DATA_BLOCK DB 50
VERSION : 0.1


  STRUCT
   STAT0 : DATE_AND_TIME  := DT#95-1-1-0:0:0.000;
   STAT1 : DATE_AND_TIME  := DT#95-1-1-0:0:0.000;
   STAT2 : INT ;
   STAT3 : DATE  := D#1995-1-1;
   STAT4 : TIME_OF_DAY ;
   STAT5 : INT ;
   STAT6 : BYTE ;
  END_STRUCT ;
BEGIN
   STAT0 := DT#22-2-18-16:13:36.401;
   STAT1 := DT#95-1-1-0:0:0.000;
   STAT2 := 0;
   STAT3 := D#1995-1-1;
   STAT4 := TOD#0:0:0.000;
   STAT5 := 0;
   STAT6 := B#16#0;
END_DATA_BLOCK

DATA_BLOCK DB 101
VERSION : 0.1


  STRUCT
   STAT0 : STRUCT
    STAT1 : STRUCT
     STAT2 : WORD ;
     STAT3 : WORD ;
    END_STRUCT ;
    STAT4 : STRUCT
     STAT5 : WORD ;
     STAT6 : STRUCT
      STAT7 : BOOL ;
      STAT8 : BOOL ;
      STAT9 : BOOL ;
      STAT10 : BOOL ;
      STAT11 : BOOL ;
      STAT12 : BOOL ;
      STAT13 : BOOL ;
      STAT14 : BOOL ;
      STAT15 : BOOL ;
      STAT16 : BOOL ;
      STAT17 : BOOL ;
      STAT18 : BOOL ;
      STAT19 : BOOL ;
      STAT20 : BOOL ;
      STAT21 : BOOL ;
      STAT22 : BOOL ;
     END_STRUCT ;
     STAT23 : WORD ;
     STAT24 : WORD ;
     STAT25 : WORD ;
     STAT26 : WORD ;
     STAT27 : WORD ;
     STAT28 : BYTE ;
     STAT29 : BYTE ;
    END_STRUCT ;
    STAT30 : BOOL ;
    STAT31 : BOOL ;
    STAT32 : WORD ;
    STAT33 : INT ;
   END_STRUCT ;
   STAT34 : STRUCT
    STAT35 : STRUCT
     STAT36 : WORD ;
     STAT37 : WORD ;
    END_STRUCT ;
    STAT38 : STRUCT
     STAT39 : ARRAY  [0 .. 12 ] OF STRUCT
      STAT40 : BOOL ;
      STAT41 : BOOL ;
      STAT42 : BOOL ;
      STAT43 : BOOL ;
      STAT44 : BOOL ;
      STAT45 : BOOL ;
      STAT46 : BOOL ;
      STAT47 : BOOL ;
      STAT48 : BYTE ;
      STAT49 : BYTE ;
      STAT50 : BYTE ;
     END_STRUCT ;
     STAT51 : ARRAY  [0 .. 12 ] OF STRUCT
      STAT52 : BOOL ;
      STAT53 : BOOL ;
      STAT54 : BOOL ;
      STAT55 : BOOL ;
      STAT56 : BOOL ;
      STAT57 : BOOL ;
      STAT58 : BOOL ;
      STAT59 : BOOL ;
      STAT60 : BYTE ;
      STAT61 : BYTE ;
      STAT62 : BYTE ;
     END_STRUCT ;
    END_STRUCT ;
    STAT63 : BOOL ;
    STAT64 : BOOL ;
    STAT65 : WORD ;
    STAT66 : INT ;
   END_STRUCT ;
   STAT67 : STRUCT
    STAT68 : STRUCT
     STAT69 : WORD ;
     STAT70 : WORD ;
    END_STRUCT ;
    STAT71 : STRUCT
     STAT72 : WORD ;
     STAT73 : WORD ;
     STAT74 : WORD ;
     STAT75 : WORD ;
     STAT76 : WORD ;
     STAT77 : WORD ;
     STAT78 : WORD ;
     STAT79 : STRUCT
      STAT80 : BOOL ;
      STAT81 : BOOL ;
      STAT82 : BOOL ;
      STAT83 : BOOL ;
      STAT84 : BOOL ;
      STAT85 : BOOL ;
      STAT86 : BOOL ;
      STAT87 : BOOL ;
      STAT88 : BOOL ;
      STAT89 : BOOL ;
      STAT90 : BOOL ;
      STAT91 : BOOL ;
      STAT92 : BOOL ;
      STAT93 : BOOL ;
      STAT94 : BOOL ;
      STAT95 : BOOL ;
     END_STRUCT ;
    END_STRUCT ;
    STAT96 : BOOL ;
    STAT97 : BOOL ;
    STAT98 : WORD ;
    STAT99 : INT ;
   END_STRUCT ;
   STAT100 : STRUCT
    STAT101 : STRUCT
     STAT102 : WORD ;
     STAT103 : WORD ;
    END_STRUCT ;
    STAT104 : STRUCT
     STAT105 : WORD ;
     STAT106 : WORD ;
     STAT107 : WORD ;
     STAT108 : WORD ;
     STAT109 : WORD ;
     STAT110 : WORD ;
     STAT111 : WORD ;
     STAT112 : STRUCT
      STAT113 : BOOL ;
      STAT114 : BOOL ;
      STAT115 : BOOL ;
      STAT116 : BOOL ;
      STAT117 : BOOL ;
      STAT118 : BOOL ;
      STAT119 : BOOL ;
      STAT120 : BOOL ;
      STAT121 : BOOL ;
      STAT122 : BOOL ;
      STAT123 : BOOL ;
      STAT124 : BOOL ;
      STAT125 : BOOL ;
      STAT126 : BOOL ;
      STAT127 : BOOL ;
      STAT128 : BOOL ;
     END_STRUCT ;
    END_STRUCT ;
    STAT129 : BOOL ;
    STAT130 : BOOL ;
    STAT131 : WORD ;
    STAT132 : INT ;
   END_STRUCT ;
   STAT133 : STRUCT
    STAT134 : STRUCT
     STAT135 : WORD ;
     STAT136 : WORD ;
    END_STRUCT ;
    STAT137 : STRUCT
     STAT138 : WORD ;
     STAT139 : WORD ;
     STAT140 : WORD ;
     STAT141 : WORD ;
     STAT142 : WORD ;
     STAT143 : WORD ;
     STAT144 : WORD ;
     STAT145 : STRUCT
      STAT146 : BOOL ;
      STAT147 : BOOL ;
      STAT148 : BOOL ;
      STAT149 : BOOL ;
      STAT150 : BOOL ;
      STAT151 : BOOL ;
      STAT152 : BOOL ;
      STAT153 : BOOL ;
      STAT154 : BOOL ;
      STAT155 : BOOL ;
      STAT156 : BOOL ;
      STAT157 : BOOL ;
      STAT158 : BOOL ;
      STAT159 : BOOL ;
      STAT160 : BOOL ;
      STAT161 : BOOL ;
     END_STRUCT ;
    END_STRUCT ;
    STAT162 : BOOL ;
    STAT163 : BOOL ;
    STAT164 : WORD ;
    STAT165 : INT ;
   END_STRUCT ;
   STAT166 : BYTE ;
   STAT167 : BYTE ;
   STAT168 : ARRAY  [0 .. 25 ] OF STRUCT
    STAT169 : BOOL ;
    STAT170 : BOOL ;
    STAT171 : BOOL ;
    STAT172 : BOOL ;
    STAT173 : BOOL ;
    STAT174 : BOOL ;
    STAT175 : BOOL ;
    STAT176 : BOOL ;
    STAT177 : BYTE ;
    STAT178 : BYTE ;
    STAT179 : BYTE ;
   END_STRUCT ;
  END_STRUCT ;
BEGIN
   STAT0.STAT1.STAT2 := W#16#10;
   STAT0.STAT1.STAT3 := W#16#1;
   STAT0.STAT4.STAT5 := W#16#12;
   STAT0.STAT4.STAT6.STAT7 := FALSE;
   STAT0.STAT4.STAT6.STAT8 := FALSE;
   STAT0.STAT4.STAT6.STAT9 := FALSE;
   STAT0.STAT4.STAT6.STAT10 := FALSE;
   STAT0.STAT4.STAT6.STAT11 := TRUE;
   STAT0.STAT4.STAT6.STAT12 := FALSE;
   STAT0.STAT4.STAT6.STAT13 := FALSE;
   STAT0.STAT4.STAT6.STAT14 := FALSE;
   STAT0.STAT4.STAT6.STAT15 := TRUE;
   STAT0.STAT4.STAT6.STAT16 := FALSE;
   STAT0.STAT4.STAT6.STAT17 := FALSE;
   STAT0.STAT4.STAT6.STAT18 := FALSE;
   STAT0.STAT4.STAT6.STAT19 := FALSE;
   STAT0.STAT4.STAT6.STAT20 := FALSE;
   STAT0.STAT4.STAT6.STAT21 := FALSE;
   STAT0.STAT4.STAT6.STAT22 := FALSE;
   STAT0.STAT4.STAT23 := W#16#0;
   STAT0.STAT4.STAT24 := W#16#0;
   STAT0.STAT4.STAT25 := W#16#9;
   STAT0.STAT4.STAT26 := W#16#9;
   STAT0.STAT4.STAT27 := W#16#0;
   STAT0.STAT4.STAT28 := B#16#3;
   STAT0.STAT4.STAT29 := B#16#0;
   STAT0.STAT30 := TRUE;
   STAT0.STAT31 := FALSE;
   STAT0.STAT32 := W#16#0;
   STAT0.STAT33 := 0;
   STAT34.STAT35.STAT36 := W#16#4;
   STAT34.STAT35.STAT37 := W#16#18;
   STAT34.STAT38.STAT39[0].STAT40 := FALSE;
   STAT34.STAT38.STAT39[0].STAT41 := FALSE;
   STAT34.STAT38.STAT39[0].STAT42 := FALSE;
   STAT34.STAT38.STAT39[0].STAT43 := TRUE;
   STAT34.STAT38.STAT39[0].STAT44 := TRUE;
   STAT34.STAT38.STAT39[0].STAT45 := TRUE;
   STAT34.STAT38.STAT39[0].STAT46 := TRUE;
   STAT34.STAT38.STAT39[0].STAT47 := TRUE;
   STAT34.STAT38.STAT39[0].STAT48 := B#16#2;
   STAT34.STAT38.STAT39[0].STAT49 := B#16#0;
   STAT34.STAT38.STAT39[0].STAT50 := B#16#0;
   STAT34.STAT38.STAT39[1].STAT40 := FALSE;
   STAT34.STAT38.STAT39[1].STAT41 := FALSE;
   STAT34.STAT38.STAT39[1].STAT42 := FALSE;
   STAT34.STAT38.STAT39[1].STAT43 := TRUE;
   STAT34.STAT38.STAT39[1].STAT44 := TRUE;
   STAT34.STAT38.STAT39[1].STAT45 := TRUE;
   STAT34.STAT38.STAT39[1].STAT46 := TRUE;
   STAT34.STAT38.STAT39[1].STAT47 := TRUE;
   STAT34.STAT38.STAT39[1].STAT48 := B#16#3;
   STAT34.STAT38.STAT39[1].STAT49 := B#16#1;
   STAT34.STAT38.STAT39[1].STAT50 := B#16#0;
   STAT34.STAT38.STAT39[2].STAT40 := FALSE;
   STAT34.STAT38.STAT39[2].STAT41 := FALSE;
   STAT34.STAT38.STAT39[2].STAT42 := FALSE;
   STAT34.STAT38.STAT39[2].STAT43 := TRUE;
   STAT34.STAT38.STAT39[2].STAT44 := TRUE;
   STAT34.STAT38.STAT39[2].STAT45 := TRUE;
   STAT34.STAT38.STAT39[2].STAT46 := TRUE;
   STAT34.STAT38.STAT39[2].STAT47 := TRUE;
   STAT34.STAT38.STAT39[2].STAT48 := B#16#4;
   STAT34.STAT38.STAT39[2].STAT49 := B#16#1;
   STAT34.STAT38.STAT39[2].STAT50 := B#16#0;
   STAT34.STAT38.STAT39[3].STAT40 := FALSE;
   STAT34.STAT38.STAT39[3].STAT41 := FALSE;
   STAT34.STAT38.STAT39[3].STAT42 := FALSE;
   STAT34.STAT38.STAT39[3].STAT43 := TRUE;
   STAT34.STAT38.STAT39[3].STAT44 := TRUE;
   STAT34.STAT38.STAT39[3].STAT45 := TRUE;
   STAT34.STAT38.STAT39[3].STAT46 := TRUE;
   STAT34.STAT38.STAT39[3].STAT47 := TRUE;
   STAT34.STAT38.STAT39[3].STAT48 := B#16#5;
   STAT34.STAT38.STAT39[3].STAT49 := B#16#0;
   STAT34.STAT38.STAT39[3].STAT50 := B#16#0;
   STAT34.STAT38.STAT39[4].STAT40 := FALSE;
   STAT34.STAT38.STAT39[4].STAT41 := FALSE;
   STAT34.STAT38.STAT39[4].STAT42 := FALSE;
   STAT34.STAT38.STAT39[4].STAT43 := TRUE;
   STAT34.STAT38.STAT39[4].STAT44 := TRUE;
   STAT34.STAT38.STAT39[4].STAT45 := TRUE;
   STAT34.STAT38.STAT39[4].STAT46 := TRUE;
   STAT34.STAT38.STAT39[4].STAT47 := TRUE;
   STAT34.STAT38.STAT39[4].STAT48 := B#16#6;
   STAT34.STAT38.STAT39[4].STAT49 := B#16#0;
   STAT34.STAT38.STAT39[4].STAT50 := B#16#0;
   STAT34.STAT38.STAT39[5].STAT40 := FALSE;
   STAT34.STAT38.STAT39[5].STAT41 := FALSE;
   STAT34.STAT38.STAT39[5].STAT42 := FALSE;
   STAT34.STAT38.STAT39[5].STAT43 := TRUE;
   STAT34.STAT38.STAT39[5].STAT44 := TRUE;
   STAT34.STAT38.STAT39[5].STAT45 := TRUE;
   STAT34.STAT38.STAT39[5].STAT46 := TRUE;
   STAT34.STAT38.STAT39[5].STAT47 := TRUE;
   STAT34.STAT38.STAT39[5].STAT48 := B#16#B;
   STAT34.STAT38.STAT39[5].STAT49 := B#16#0;
   STAT34.STAT38.STAT39[5].STAT50 := B#16#0;
   STAT34.STAT38.STAT39[6].STAT40 := FALSE;
   STAT34.STAT38.STAT39[6].STAT41 := FALSE;
   STAT34.STAT38.STAT39[6].STAT42 := FALSE;
   STAT34.STAT38.STAT39[6].STAT43 := TRUE;
   STAT34.STAT38.STAT39[6].STAT44 := TRUE;
   STAT34.STAT38.STAT39[6].STAT45 := TRUE;
   STAT34.STAT38.STAT39[6].STAT46 := TRUE;
   STAT34.STAT38.STAT39[6].STAT47 := TRUE;
   STAT34.STAT38.STAT39[6].STAT48 := B#16#D;
   STAT34.STAT38.STAT39[6].STAT49 := B#16#0;
   STAT34.STAT38.STAT39[6].STAT50 := B#16#0;
   STAT34.STAT38.STAT39[7].STAT40 := FALSE;
   STAT34.STAT38.STAT39[7].STAT41 := FALSE;
   STAT34.STAT38.STAT39[7].STAT42 := FALSE;
   STAT34.STAT38.STAT39[7].STAT43 := TRUE;
   STAT34.STAT38.STAT39[7].STAT44 := TRUE;
   STAT34.STAT38.STAT39[7].STAT45 := TRUE;
   STAT34.STAT38.STAT39[7].STAT46 := TRUE;
   STAT34.STAT38.STAT39[7].STAT47 := TRUE;
   STAT34.STAT38.STAT39[7].STAT48 := B#16#E;
   STAT34.STAT38.STAT39[7].STAT49 := B#16#1;
   STAT34.STAT38.STAT39[7].STAT50 := B#16#0;
   STAT34.STAT38.STAT39[8].STAT40 := FALSE;
   STAT34.STAT38.STAT39[8].STAT41 := FALSE;
   STAT34.STAT38.STAT39[8].STAT42 := FALSE;
   STAT34.STAT38.STAT39[8].STAT43 := TRUE;
   STAT34.STAT38.STAT39[8].STAT44 := TRUE;
   STAT34.STAT38.STAT39[8].STAT45 := TRUE;
   STAT34.STAT38.STAT39[8].STAT46 := TRUE;
   STAT34.STAT38.STAT39[8].STAT47 := TRUE;
   STAT34.STAT38.STAT39[8].STAT48 := B#16#F;
   STAT34.STAT38.STAT39[8].STAT49 := B#16#1;
   STAT34.STAT38.STAT39[8].STAT50 := B#16#0;
   STAT34.STAT38.STAT39[9].STAT40 := FALSE;
   STAT34.STAT38.STAT39[9].STAT41 := FALSE;
   STAT34.STAT38.STAT39[9].STAT42 := FALSE;
   STAT34.STAT38.STAT39[9].STAT43 := TRUE;
   STAT34.STAT38.STAT39[9].STAT44 := TRUE;
   STAT34.STAT38.STAT39[9].STAT45 := TRUE;
   STAT34.STAT38.STAT39[9].STAT46 := TRUE;
   STAT34.STAT38.STAT39[9].STAT47 := TRUE;
   STAT34.STAT38.STAT39[9].STAT48 := B#16#10;
   STAT34.STAT38.STAT39[9].STAT49 := B#16#0;
   STAT34.STAT38.STAT39[9].STAT50 := B#16#0;
   STAT34.STAT38.STAT39[10].STAT40 := FALSE;
   STAT34.STAT38.STAT39[10].STAT41 := FALSE;
   STAT34.STAT38.STAT39[10].STAT42 := FALSE;
   STAT34.STAT38.STAT39[10].STAT43 := TRUE;
   STAT34.STAT38.STAT39[10].STAT44 := TRUE;
   STAT34.STAT38.STAT39[10].STAT45 := TRUE;
   STAT34.STAT38.STAT39[10].STAT46 := TRUE;
   STAT34.STAT38.STAT39[10].STAT47 := TRUE;
   STAT34.STAT38.STAT39[10].STAT48 := B#16#12;
   STAT34.STAT38.STAT39[10].STAT49 := B#16#0;
   STAT34.STAT38.STAT39[10].STAT50 := B#16#0;
   STAT34.STAT38.STAT39[11].STAT40 := FALSE;
   STAT34.STAT38.STAT39[11].STAT41 := FALSE;
   STAT34.STAT38.STAT39[11].STAT42 := FALSE;
   STAT34.STAT38.STAT39[11].STAT43 := TRUE;
   STAT34.STAT38.STAT39[11].STAT44 := TRUE;
   STAT34.STAT38.STAT39[11].STAT45 := TRUE;
   STAT34.STAT38.STAT39[11].STAT46 := TRUE;
   STAT34.STAT38.STAT39[11].STAT47 := TRUE;
   STAT34.STAT38.STAT39[11].STAT48 := B#16#13;
   STAT34.STAT38.STAT39[11].STAT49 := B#16#0;
   STAT34.STAT38.STAT39[11].STAT50 := B#16#0;
   STAT34.STAT38.STAT39[12].STAT40 := TRUE;
   STAT34.STAT38.STAT39[12].STAT41 := FALSE;
   STAT34.STAT38.STAT39[12].STAT42 := FALSE;
   STAT34.STAT38.STAT39[12].STAT43 := FALSE;
   STAT34.STAT38.STAT39[12].STAT44 := TRUE;
   STAT34.STAT38.STAT39[12].STAT45 := TRUE;
   STAT34.STAT38.STAT39[12].STAT46 := TRUE;
   STAT34.STAT38.STAT39[12].STAT47 := TRUE;
   STAT34.STAT38.STAT39[12].STAT48 := B#16#2;
   STAT34.STAT38.STAT39[12].STAT49 := B#16#0;
   STAT34.STAT38.STAT39[12].STAT50 := B#16#0;
   STAT34.STAT38.STAT51[0].STAT52 := TRUE;
   STAT34.STAT38.STAT51[0].STAT53 := FALSE;
   STAT34.STAT38.STAT51[0].STAT54 := FALSE;
   STAT34.STAT38.STAT51[0].STAT55 := FALSE;
   STAT34.STAT38.STAT51[0].STAT56 := TRUE;
   STAT34.STAT38.STAT51[0].STAT57 := TRUE;
   STAT34.STAT38.STAT51[0].STAT58 := TRUE;
   STAT34.STAT38.STAT51[0].STAT59 := TRUE;
   STAT34.STAT38.STAT51[0].STAT60 := B#16#3;
   STAT34.STAT38.STAT51[0].STAT61 := B#16#1;
   STAT34.STAT38.STAT51[0].STAT62 := B#16#0;
   STAT34.STAT38.STAT51[1].STAT52 := TRUE;
   STAT34.STAT38.STAT51[1].STAT53 := FALSE;
   STAT34.STAT38.STAT51[1].STAT54 := FALSE;
   STAT34.STAT38.STAT51[1].STAT55 := FALSE;
   STAT34.STAT38.STAT51[1].STAT56 := TRUE;
   STAT34.STAT38.STAT51[1].STAT57 := TRUE;
   STAT34.STAT38.STAT51[1].STAT58 := TRUE;
   STAT34.STAT38.STAT51[1].STAT59 := TRUE;
   STAT34.STAT38.STAT51[1].STAT60 := B#16#4;
   STAT34.STAT38.STAT51[1].STAT61 := B#16#1;
   STAT34.STAT38.STAT51[1].STAT62 := B#16#0;
   STAT34.STAT38.STAT51[2].STAT52 := TRUE;
   STAT34.STAT38.STAT51[2].STAT53 := FALSE;
   STAT34.STAT38.STAT51[2].STAT54 := FALSE;
   STAT34.STAT38.STAT51[2].STAT55 := FALSE;
   STAT34.STAT38.STAT51[2].STAT56 := TRUE;
   STAT34.STAT38.STAT51[2].STAT57 := TRUE;
   STAT34.STAT38.STAT51[2].STAT58 := TRUE;
   STAT34.STAT38.STAT51[2].STAT59 := TRUE;
   STAT34.STAT38.STAT51[2].STAT60 := B#16#5;
   STAT34.STAT38.STAT51[2].STAT61 := B#16#0;
   STAT34.STAT38.STAT51[2].STAT62 := B#16#0;
   STAT34.STAT38.STAT51[3].STAT52 := TRUE;
   STAT34.STAT38.STAT51[3].STAT53 := FALSE;
   STAT34.STAT38.STAT51[3].STAT54 := FALSE;
   STAT34.STAT38.STAT51[3].STAT55 := FALSE;
   STAT34.STAT38.STAT51[3].STAT56 := TRUE;
   STAT34.STAT38.STAT51[3].STAT57 := TRUE;
   STAT34.STAT38.STAT51[3].STAT58 := TRUE;
   STAT34.STAT38.STAT51[3].STAT59 := TRUE;
   STAT34.STAT38.STAT51[3].STAT60 := B#16#6;
   STAT34.STAT38.STAT51[3].STAT61 := B#16#0;
   STAT34.STAT38.STAT51[3].STAT62 := B#16#0;
   STAT34.STAT38.STAT51[4].STAT52 := TRUE;
   STAT34.STAT38.STAT51[4].STAT53 := FALSE;
   STAT34.STAT38.STAT51[4].STAT54 := FALSE;
   STAT34.STAT38.STAT51[4].STAT55 := FALSE;
   STAT34.STAT38.STAT51[4].STAT56 := TRUE;
   STAT34.STAT38.STAT51[4].STAT57 := TRUE;
   STAT34.STAT38.STAT51[4].STAT58 := TRUE;
   STAT34.STAT38.STAT51[4].STAT59 := TRUE;
   STAT34.STAT38.STAT51[4].STAT60 := B#16#B;
   STAT34.STAT38.STAT51[4].STAT61 := B#16#0;
   STAT34.STAT38.STAT51[4].STAT62 := B#16#0;
   STAT34.STAT38.STAT51[5].STAT52 := TRUE;
   STAT34.STAT38.STAT51[5].STAT53 := FALSE;
   STAT34.STAT38.STAT51[5].STAT54 := FALSE;
   STAT34.STAT38.STAT51[5].STAT55 := FALSE;
   STAT34.STAT38.STAT51[5].STAT56 := TRUE;
   STAT34.STAT38.STAT51[5].STAT57 := TRUE;
   STAT34.STAT38.STAT51[5].STAT58 := TRUE;
   STAT34.STAT38.STAT51[5].STAT59 := TRUE;
   STAT34.STAT38.STAT51[5].STAT60 := B#16#D;
   STAT34.STAT38.STAT51[5].STAT61 := B#16#0;
   STAT34.STAT38.STAT51[5].STAT62 := B#16#0;
   STAT34.STAT38.STAT51[6].STAT52 := TRUE;
   STAT34.STAT38.STAT51[6].STAT53 := FALSE;
   STAT34.STAT38.STAT51[6].STAT54 := FALSE;
   STAT34.STAT38.STAT51[6].STAT55 := FALSE;
   STAT34.STAT38.STAT51[6].STAT56 := TRUE;
   STAT34.STAT38.STAT51[6].STAT57 := TRUE;
   STAT34.STAT38.STAT51[6].STAT58 := TRUE;
   STAT34.STAT38.STAT51[6].STAT59 := TRUE;
   STAT34.STAT38.STAT51[6].STAT60 := B#16#E;
   STAT34.STAT38.STAT51[6].STAT61 := B#16#0;
   STAT34.STAT38.STAT51[6].STAT62 := B#16#0;
   STAT34.STAT38.STAT51[7].STAT52 := TRUE;
   STAT34.STAT38.STAT51[7].STAT53 := FALSE;
   STAT34.STAT38.STAT51[7].STAT54 := FALSE;
   STAT34.STAT38.STAT51[7].STAT55 := FALSE;
   STAT34.STAT38.STAT51[7].STAT56 := TRUE;
   STAT34.STAT38.STAT51[7].STAT57 := TRUE;
   STAT34.STAT38.STAT51[7].STAT58 := TRUE;
   STAT34.STAT38.STAT51[7].STAT59 := TRUE;
   STAT34.STAT38.STAT51[7].STAT60 := B#16#F;
   STAT34.STAT38.STAT51[7].STAT61 := B#16#0;
   STAT34.STAT38.STAT51[7].STAT62 := B#16#0;
   STAT34.STAT38.STAT51[8].STAT52 := TRUE;
   STAT34.STAT38.STAT51[8].STAT53 := FALSE;
   STAT34.STAT38.STAT51[8].STAT54 := FALSE;
   STAT34.STAT38.STAT51[8].STAT55 := FALSE;
   STAT34.STAT38.STAT51[8].STAT56 := TRUE;
   STAT34.STAT38.STAT51[8].STAT57 := TRUE;
   STAT34.STAT38.STAT51[8].STAT58 := TRUE;
   STAT34.STAT38.STAT51[8].STAT59 := TRUE;
   STAT34.STAT38.STAT51[8].STAT60 := B#16#10;
   STAT34.STAT38.STAT51[8].STAT61 := B#16#1;
   STAT34.STAT38.STAT51[8].STAT62 := B#16#0;
   STAT34.STAT38.STAT51[9].STAT52 := TRUE;
   STAT34.STAT38.STAT51[9].STAT53 := FALSE;
   STAT34.STAT38.STAT51[9].STAT54 := FALSE;
   STAT34.STAT38.STAT51[9].STAT55 := FALSE;
   STAT34.STAT38.STAT51[9].STAT56 := TRUE;
   STAT34.STAT38.STAT51[9].STAT57 := TRUE;
   STAT34.STAT38.STAT51[9].STAT58 := TRUE;
   STAT34.STAT38.STAT51[9].STAT59 := TRUE;
   STAT34.STAT38.STAT51[9].STAT60 := B#16#12;
   STAT34.STAT38.STAT51[9].STAT61 := B#16#0;
   STAT34.STAT38.STAT51[9].STAT62 := B#16#0;
   STAT34.STAT38.STAT51[10].STAT52 := TRUE;
   STAT34.STAT38.STAT51[10].STAT53 := FALSE;
   STAT34.STAT38.STAT51[10].STAT54 := FALSE;
   STAT34.STAT38.STAT51[10].STAT55 := FALSE;
   STAT34.STAT38.STAT51[10].STAT56 := TRUE;
   STAT34.STAT38.STAT51[10].STAT57 := TRUE;
   STAT34.STAT38.STAT51[10].STAT58 := TRUE;
   STAT34.STAT38.STAT51[10].STAT59 := TRUE;
   STAT34.STAT38.STAT51[10].STAT60 := B#16#13;
   STAT34.STAT38.STAT51[10].STAT61 := B#16#0;
   STAT34.STAT38.STAT51[10].STAT62 := B#16#0;
   STAT34.STAT38.STAT51[11].STAT52 := FALSE;
   STAT34.STAT38.STAT51[11].STAT53 := FALSE;
   STAT34.STAT38.STAT51[11].STAT54 := FALSE;
   STAT34.STAT38.STAT51[11].STAT55 := FALSE;
   STAT34.STAT38.STAT51[11].STAT56 := FALSE;
   STAT34.STAT38.STAT51[11].STAT57 := FALSE;
   STAT34.STAT38.STAT51[11].STAT58 := FALSE;
   STAT34.STAT38.STAT51[11].STAT59 := FALSE;
   STAT34.STAT38.STAT51[11].STAT60 := B#16#0;
   STAT34.STAT38.STAT51[11].STAT61 := B#16#0;
   STAT34.STAT38.STAT51[11].STAT62 := B#16#0;
   STAT34.STAT38.STAT51[12].STAT52 := FALSE;
   STAT34.STAT38.STAT51[12].STAT53 := FALSE;
   STAT34.STAT38.STAT51[12].STAT54 := FALSE;
   STAT34.STAT38.STAT51[12].STAT55 := FALSE;
   STAT34.STAT38.STAT51[12].STAT56 := FALSE;
   STAT34.STAT38.STAT51[12].STAT57 := FALSE;
   STAT34.STAT38.STAT51[12].STAT58 := FALSE;
   STAT34.STAT38.STAT51[12].STAT59 := FALSE;
   STAT34.STAT38.STAT51[12].STAT60 := B#16#0;
   STAT34.STAT38.STAT51[12].STAT61 := B#16#0;
   STAT34.STAT38.STAT51[12].STAT62 := B#16#0;
   STAT34.STAT63 := TRUE;
   STAT34.STAT64 := FALSE;
   STAT34.STAT65 := W#16#0;
   STAT34.STAT66 := 0;
   STAT67.STAT68.STAT69 := W#16#0;
   STAT67.STAT68.STAT70 := W#16#0;
   STAT67.STAT71.STAT72 := W#16#0;
   STAT67.STAT71.STAT73 := W#16#0;
   STAT67.STAT71.STAT74 := W#16#0;
   STAT67.STAT71.STAT75 := W#16#0;
   STAT67.STAT71.STAT76 := W#16#0;
   STAT67.STAT71.STAT77 := W#16#0;
   STAT67.STAT71.STAT78 := W#16#0;
   STAT67.STAT71.STAT79.STAT80 := FALSE;
   STAT67.STAT71.STAT79.STAT81 := FALSE;
   STAT67.STAT71.STAT79.STAT82 := FALSE;
   STAT67.STAT71.STAT79.STAT83 := FALSE;
   STAT67.STAT71.STAT79.STAT84 := FALSE;
   STAT67.STAT71.STAT79.STAT85 := FALSE;
   STAT67.STAT71.STAT79.STAT86 := FALSE;
   STAT67.STAT71.STAT79.STAT87 := FALSE;
   STAT67.STAT71.STAT79.STAT88 := FALSE;
   STAT67.STAT71.STAT79.STAT89 := FALSE;
   STAT67.STAT71.STAT79.STAT90 := FALSE;
   STAT67.STAT71.STAT79.STAT91 := FALSE;
   STAT67.STAT71.STAT79.STAT92 := FALSE;
   STAT67.STAT71.STAT79.STAT93 := FALSE;
   STAT67.STAT71.STAT79.STAT94 := FALSE;
   STAT67.STAT71.STAT79.STAT95 := FALSE;
   STAT67.STAT96 := FALSE;
   STAT67.STAT97 := FALSE;
   STAT67.STAT98 := W#16#0;
   STAT67.STAT99 := 0;
   STAT100.STAT101.STAT102 := W#16#0;
   STAT100.STAT101.STAT103 := W#16#0;
   STAT100.STAT104.STAT105 := W#16#0;
   STAT100.STAT104.STAT106 := W#16#0;
   STAT100.STAT104.STAT107 := W#16#0;
   STAT100.STAT104.STAT108 := W#16#0;
   STAT100.STAT104.STAT109 := W#16#0;
   STAT100.STAT104.STAT110 := W#16#0;
   STAT100.STAT104.STAT111 := W#16#0;
   STAT100.STAT104.STAT112.STAT113 := FALSE;
   STAT100.STAT104.STAT112.STAT114 := FALSE;
   STAT100.STAT104.STAT112.STAT115 := FALSE;
   STAT100.STAT104.STAT112.STAT116 := FALSE;
   STAT100.STAT104.STAT112.STAT117 := FALSE;
   STAT100.STAT104.STAT112.STAT118 := FALSE;
   STAT100.STAT104.STAT112.STAT119 := FALSE;
   STAT100.STAT104.STAT112.STAT120 := FALSE;
   STAT100.STAT104.STAT112.STAT121 := FALSE;
   STAT100.STAT104.STAT112.STAT122 := FALSE;
   STAT100.STAT104.STAT112.STAT123 := FALSE;
   STAT100.STAT104.STAT112.STAT124 := FALSE;
   STAT100.STAT104.STAT112.STAT125 := FALSE;
   STAT100.STAT104.STAT112.STAT126 := FALSE;
   STAT100.STAT104.STAT112.STAT127 := FALSE;
   STAT100.STAT104.STAT112.STAT128 := FALSE;
   STAT100.STAT129 := FALSE;
   STAT100.STAT130 := FALSE;
   STAT100.STAT131 := W#16#0;
   STAT100.STAT132 := 0;
   STAT133.STAT134.STAT135 := W#16#0;
   STAT133.STAT134.STAT136 := W#16#0;
   STAT133.STAT137.STAT138 := W#16#0;
   STAT133.STAT137.STAT139 := W#16#0;
   STAT133.STAT137.STAT140 := W#16#0;
   STAT133.STAT137.STAT141 := W#16#0;
   STAT133.STAT137.STAT142 := W#16#0;
   STAT133.STAT137.STAT143 := W#16#0;
   STAT133.STAT137.STAT144 := W#16#0;
   STAT133.STAT137.STAT145.STAT146 := FALSE;
   STAT133.STAT137.STAT145.STAT147 := FALSE;
   STAT133.STAT137.STAT145.STAT148 := FALSE;
   STAT133.STAT137.STAT145.STAT149 := FALSE;
   STAT133.STAT137.STAT145.STAT150 := FALSE;
   STAT133.STAT137.STAT145.STAT151 := FALSE;
   STAT133.STAT137.STAT145.STAT152 := FALSE;
   STAT133.STAT137.STAT145.STAT153 := FALSE;
   STAT133.STAT137.STAT145.STAT154 := FALSE;
   STAT133.STAT137.STAT145.STAT155 := FALSE;
   STAT133.STAT137.STAT145.STAT156 := FALSE;
   STAT133.STAT137.STAT145.STAT157 := FALSE;
   STAT133.STAT137.STAT145.STAT158 := FALSE;
   STAT133.STAT137.STAT145.STAT159 := FALSE;
   STAT133.STAT137.STAT145.STAT160 := FALSE;
   STAT133.STAT137.STAT145.STAT161 := FALSE;
   STAT133.STAT162 := FALSE;
   STAT133.STAT163 := FALSE;
   STAT133.STAT164 := W#16#0;
   STAT133.STAT165 := 0;
   STAT166 := B#16#0;
   STAT167 := B#16#0;
   STAT168[0].STAT169 := FALSE;
   STAT168[0].STAT170 := FALSE;
   STAT168[0].STAT171 := FALSE;
   STAT168[0].STAT172 := FALSE;
   STAT168[0].STAT173 := FALSE;
   STAT168[0].STAT174 := FALSE;
   STAT168[0].STAT175 := FALSE;
   STAT168[0].STAT176 := FALSE;
   STAT168[0].STAT177 := B#16#0;
   STAT168[0].STAT178 := B#16#0;
   STAT168[0].STAT179 := B#16#0;
   STAT168[1].STAT169 := FALSE;
   STAT168[1].STAT170 := FALSE;
   STAT168[1].STAT171 := FALSE;
   STAT168[1].STAT172 := FALSE;
   STAT168[1].STAT173 := FALSE;
   STAT168[1].STAT174 := FALSE;
   STAT168[1].STAT175 := FALSE;
   STAT168[1].STAT176 := FALSE;
   STAT168[1].STAT177 := B#16#0;
   STAT168[1].STAT178 := B#16#0;
   STAT168[1].STAT179 := B#16#0;
   STAT168[2].STAT169 := FALSE;
   STAT168[2].STAT170 := FALSE;
   STAT168[2].STAT171 := FALSE;
   STAT168[2].STAT172 := FALSE;
   STAT168[2].STAT173 := FALSE;
   STAT168[2].STAT174 := FALSE;
   STAT168[2].STAT175 := FALSE;
   STAT168[2].STAT176 := FALSE;
   STAT168[2].STAT177 := B#16#0;
   STAT168[2].STAT178 := B#16#0;
   STAT168[2].STAT179 := B#16#0;
   STAT168[3].STAT169 := FALSE;
   STAT168[3].STAT170 := FALSE;
   STAT168[3].STAT171 := FALSE;
   STAT168[3].STAT172 := FALSE;
   STAT168[3].STAT173 := FALSE;
   STAT168[3].STAT174 := FALSE;
   STAT168[3].STAT175 := FALSE;
   STAT168[3].STAT176 := FALSE;
   STAT168[3].STAT177 := B#16#0;
   STAT168[3].STAT178 := B#16#0;
   STAT168[3].STAT179 := B#16#0;
   STAT168[4].STAT169 := FALSE;
   STAT168[4].STAT170 := FALSE;
   STAT168[4].STAT171 := FALSE;
   STAT168[4].STAT172 := FALSE;
   STAT168[4].STAT173 := FALSE;
   STAT168[4].STAT174 := FALSE;
   STAT168[4].STAT175 := FALSE;
   STAT168[4].STAT176 := FALSE;
   STAT168[4].STAT177 := B#16#0;
   STAT168[4].STAT178 := B#16#0;
   STAT168[4].STAT179 := B#16#0;
   STAT168[5].STAT169 := FALSE;
   STAT168[5].STAT170 := FALSE;
   STAT168[5].STAT171 := FALSE;
   STAT168[5].STAT172 := FALSE;
   STAT168[5].STAT173 := FALSE;
   STAT168[5].STAT174 := FALSE;
   STAT168[5].STAT175 := FALSE;
   STAT168[5].STAT176 := FALSE;
   STAT168[5].STAT177 := B#16#0;
   STAT168[5].STAT178 := B#16#0;
   STAT168[5].STAT179 := B#16#0;
   STAT168[6].STAT169 := FALSE;
   STAT168[6].STAT170 := FALSE;
   STAT168[6].STAT171 := FALSE;
   STAT168[6].STAT172 := FALSE;
   STAT168[6].STAT173 := FALSE;
   STAT168[6].STAT174 := FALSE;
   STAT168[6].STAT175 := FALSE;
   STAT168[6].STAT176 := FALSE;
   STAT168[6].STAT177 := B#16#0;
   STAT168[6].STAT178 := B#16#0;
   STAT168[6].STAT179 := B#16#0;
   STAT168[7].STAT169 := FALSE;
   STAT168[7].STAT170 := FALSE;
   STAT168[7].STAT171 := FALSE;
   STAT168[7].STAT172 := FALSE;
   STAT168[7].STAT173 := FALSE;
   STAT168[7].STAT174 := FALSE;
   STAT168[7].STAT175 := FALSE;
   STAT168[7].STAT176 := FALSE;
   STAT168[7].STAT177 := B#16#0;
   STAT168[7].STAT178 := B#16#0;
   STAT168[7].STAT179 := B#16#0;
   STAT168[8].STAT169 := FALSE;
   STAT168[8].STAT170 := FALSE;
   STAT168[8].STAT171 := FALSE;
   STAT168[8].STAT172 := FALSE;
   STAT168[8].STAT173 := FALSE;
   STAT168[8].STAT174 := FALSE;
   STAT168[8].STAT175 := FALSE;
   STAT168[8].STAT176 := FALSE;
   STAT168[8].STAT177 := B#16#0;
   STAT168[8].STAT178 := B#16#0;
   STAT168[8].STAT179 := B#16#0;
   STAT168[9].STAT169 := FALSE;
   STAT168[9].STAT170 := FALSE;
   STAT168[9].STAT171 := FALSE;
   STAT168[9].STAT172 := FALSE;
   STAT168[9].STAT173 := FALSE;
   STAT168[9].STAT174 := FALSE;
   STAT168[9].STAT175 := FALSE;
   STAT168[9].STAT176 := FALSE;
   STAT168[9].STAT177 := B#16#0;
   STAT168[9].STAT178 := B#16#0;
   STAT168[9].STAT179 := B#16#0;
   STAT168[10].STAT169 := FALSE;
   STAT168[10].STAT170 := FALSE;
   STAT168[10].STAT171 := FALSE;
   STAT168[10].STAT172 := FALSE;
   STAT168[10].STAT173 := FALSE;
   STAT168[10].STAT174 := FALSE;
   STAT168[10].STAT175 := FALSE;
   STAT168[10].STAT176 := FALSE;
   STAT168[10].STAT177 := B#16#0;
   STAT168[10].STAT178 := B#16#0;
   STAT168[10].STAT179 := B#16#0;
   STAT168[11].STAT169 := FALSE;
   STAT168[11].STAT170 := FALSE;
   STAT168[11].STAT171 := FALSE;
   STAT168[11].STAT172 := FALSE;
   STAT168[11].STAT173 := FALSE;
   STAT168[11].STAT174 := FALSE;
   STAT168[11].STAT175 := FALSE;
   STAT168[11].STAT176 := FALSE;
   STAT168[11].STAT177 := B#16#0;
   STAT168[11].STAT178 := B#16#0;
   STAT168[11].STAT179 := B#16#0;
   STAT168[12].STAT169 := FALSE;
   STAT168[12].STAT170 := FALSE;
   STAT168[12].STAT171 := FALSE;
   STAT168[12].STAT172 := FALSE;
   STAT168[12].STAT173 := FALSE;
   STAT168[12].STAT174 := FALSE;
   STAT168[12].STAT175 := FALSE;
   STAT168[12].STAT176 := FALSE;
   STAT168[12].STAT177 := B#16#0;
   STAT168[12].STAT178 := B#16#0;
   STAT168[12].STAT179 := B#16#0;
   STAT168[13].STAT169 := FALSE;
   STAT168[13].STAT170 := FALSE;
   STAT168[13].STAT171 := FALSE;
   STAT168[13].STAT172 := FALSE;
   STAT168[13].STAT173 := FALSE;
   STAT168[13].STAT174 := FALSE;
   STAT168[13].STAT175 := FALSE;
   STAT168[13].STAT176 := FALSE;
   STAT168[13].STAT177 := B#16#0;
   STAT168[13].STAT178 := B#16#0;
   STAT168[13].STAT179 := B#16#0;
   STAT168[14].STAT169 := FALSE;
   STAT168[14].STAT170 := FALSE;
   STAT168[14].STAT171 := FALSE;
   STAT168[14].STAT172 := FALSE;
   STAT168[14].STAT173 := FALSE;
   STAT168[14].STAT174 := FALSE;
   STAT168[14].STAT175 := FALSE;
   STAT168[14].STAT176 := FALSE;
   STAT168[14].STAT177 := B#16#0;
   STAT168[14].STAT178 := B#16#0;
   STAT168[14].STAT179 := B#16#0;
   STAT168[15].STAT169 := FALSE;
   STAT168[15].STAT170 := FALSE;
   STAT168[15].STAT171 := FALSE;
   STAT168[15].STAT172 := FALSE;
   STAT168[15].STAT173 := FALSE;
   STAT168[15].STAT174 := FALSE;
   STAT168[15].STAT175 := FALSE;
   STAT168[15].STAT176 := FALSE;
   STAT168[15].STAT177 := B#16#0;
   STAT168[15].STAT178 := B#16#0;
   STAT168[15].STAT179 := B#16#0;
   STAT168[16].STAT169 := FALSE;
   STAT168[16].STAT170 := FALSE;
   STAT168[16].STAT171 := FALSE;
   STAT168[16].STAT172 := FALSE;
   STAT168[16].STAT173 := FALSE;
   STAT168[16].STAT174 := FALSE;
   STAT168[16].STAT175 := FALSE;
   STAT168[16].STAT176 := FALSE;
   STAT168[16].STAT177 := B#16#0;
   STAT168[16].STAT178 := B#16#0;
   STAT168[16].STAT179 := B#16#0;
   STAT168[17].STAT169 := FALSE;
   STAT168[17].STAT170 := FALSE;
   STAT168[17].STAT171 := FALSE;
   STAT168[17].STAT172 := FALSE;
   STAT168[17].STAT173 := FALSE;
   STAT168[17].STAT174 := FALSE;
   STAT168[17].STAT175 := FALSE;
   STAT168[17].STAT176 := FALSE;
   STAT168[17].STAT177 := B#16#0;
   STAT168[17].STAT178 := B#16#0;
   STAT168[17].STAT179 := B#16#0;
   STAT168[18].STAT169 := FALSE;
   STAT168[18].STAT170 := FALSE;
   STAT168[18].STAT171 := FALSE;
   STAT168[18].STAT172 := FALSE;
   STAT168[18].STAT173 := FALSE;
   STAT168[18].STAT174 := FALSE;
   STAT168[18].STAT175 := FALSE;
   STAT168[18].STAT176 := FALSE;
   STAT168[18].STAT177 := B#16#0;
   STAT168[18].STAT178 := B#16#0;
   STAT168[18].STAT179 := B#16#0;
   STAT168[19].STAT169 := FALSE;
   STAT168[19].STAT170 := FALSE;
   STAT168[19].STAT171 := FALSE;
   STAT168[19].STAT172 := FALSE;
   STAT168[19].STAT173 := FALSE;
   STAT168[19].STAT174 := FALSE;
   STAT168[19].STAT175 := FALSE;
   STAT168[19].STAT176 := FALSE;
   STAT168[19].STAT177 := B#16#0;
   STAT168[19].STAT178 := B#16#0;
   STAT168[19].STAT179 := B#16#0;
   STAT168[20].STAT169 := FALSE;
   STAT168[20].STAT170 := FALSE;
   STAT168[20].STAT171 := FALSE;
   STAT168[20].STAT172 := FALSE;
   STAT168[20].STAT173 := FALSE;
   STAT168[20].STAT174 := FALSE;
   STAT168[20].STAT175 := FALSE;
   STAT168[20].STAT176 := FALSE;
   STAT168[20].STAT177 := B#16#0;
   STAT168[20].STAT178 := B#16#0;
   STAT168[20].STAT179 := B#16#0;
   STAT168[21].STAT169 := FALSE;
   STAT168[21].STAT170 := FALSE;
   STAT168[21].STAT171 := FALSE;
   STAT168[21].STAT172 := FALSE;
   STAT168[21].STAT173 := FALSE;
   STAT168[21].STAT174 := FALSE;
   STAT168[21].STAT175 := FALSE;
   STAT168[21].STAT176 := FALSE;
   STAT168[21].STAT177 := B#16#0;
   STAT168[21].STAT178 := B#16#0;
   STAT168[21].STAT179 := B#16#0;
   STAT168[22].STAT169 := FALSE;
   STAT168[22].STAT170 := FALSE;
   STAT168[22].STAT171 := FALSE;
   STAT168[22].STAT172 := FALSE;
   STAT168[22].STAT173 := FALSE;
   STAT168[22].STAT174 := FALSE;
   STAT168[22].STAT175 := FALSE;
   STAT168[22].STAT176 := FALSE;
   STAT168[22].STAT177 := B#16#0;
   STAT168[22].STAT178 := B#16#0;
   STAT168[22].STAT179 := B#16#0;
   STAT168[23].STAT169 := FALSE;
   STAT168[23].STAT170 := FALSE;
   STAT168[23].STAT171 := FALSE;
   STAT168[23].STAT172 := FALSE;
   STAT168[23].STAT173 := FALSE;
   STAT168[23].STAT174 := FALSE;
   STAT168[23].STAT175 := FALSE;
   STAT168[23].STAT176 := FALSE;
   STAT168[23].STAT177 := B#16#0;
   STAT168[23].STAT178 := B#16#0;
   STAT168[23].STAT179 := B#16#0;
   STAT168[24].STAT169 := FALSE;
   STAT168[24].STAT170 := FALSE;
   STAT168[24].STAT171 := FALSE;
   STAT168[24].STAT172 := FALSE;
   STAT168[24].STAT173 := FALSE;
   STAT168[24].STAT174 := FALSE;
   STAT168[24].STAT175 := FALSE;
   STAT168[24].STAT176 := FALSE;
   STAT168[24].STAT177 := B#16#0;
   STAT168[24].STAT178 := B#16#0;
   STAT168[24].STAT179 := B#16#0;
   STAT168[25].STAT169 := FALSE;
   STAT168[25].STAT170 := FALSE;
   STAT168[25].STAT171 := FALSE;
   STAT168[25].STAT172 := FALSE;
   STAT168[25].STAT173 := FALSE;
   STAT168[25].STAT174 := FALSE;
   STAT168[25].STAT175 := FALSE;
   STAT168[25].STAT176 := FALSE;
   STAT168[25].STAT177 := B#16#0;
   STAT168[25].STAT178 := B#16#0;
   STAT168[25].STAT179 := B#16#0;
END_DATA_BLOCK

DATA_BLOCK DB 103
VERSION : 0.1


  STRUCT
   STAT0 : BOOL ;
   STAT1 : BOOL ;
   STAT2 : BOOL ;
   STAT3 : WORD ;
   STAT4 : INT ;
   STAT5 : STRUCT
    STAT6 : BYTE ;
    STAT7 : BYTE ;
    STAT8 : BYTE ;
    STAT9 : BYTE ;
    STAT10 : BYTE ;
    STAT11 : BYTE ;
    STAT12 : BYTE ;
    STAT13 : BYTE ;
    STAT14 : BYTE ;
    STAT15 : BYTE ;
    STAT16 : ARRAY  [0 .. 230 ] OF BYTE ;
   END_STRUCT ;
  END_STRUCT ;
BEGIN
   STAT0 := TRUE;
   STAT1 := FALSE;
   STAT2 := FALSE;
   STAT3 := W#16#1FF7;
   STAT4 := 25;
   STAT5.STAT6 := B#16#0;
   STAT5.STAT7 := B#16#C;
   STAT5.STAT8 := B#16#0;
   STAT5.STAT9 := B#16#2;
   STAT5.STAT10 := B#16#80;
   STAT5.STAT11 := B#16#1E;
   STAT5.STAT12 := B#16#43;
   STAT5.STAT13 := B#16#0;
   STAT5.STAT14 := B#16#0;
   STAT5.STAT15 := B#16#8;
   STAT5.STAT16[0] := B#16#82;
   STAT5.STAT16[1] := B#16#0;
   STAT5.STAT16[2] := B#16#0;
   STAT5.STAT16[3] := B#16#0;
   STAT5.STAT16[4] := B#16#0;
   STAT5.STAT16[5] := B#16#0;
   STAT5.STAT16[6] := B#16#0;
   STAT5.STAT16[7] := B#16#8;
   STAT5.STAT16[8] := B#16#9F;
   STAT5.STAT16[9] := B#16#0;
   STAT5.STAT16[10] := B#16#C8;
   STAT5.STAT16[11] := B#16#42;
   STAT5.STAT16[12] := B#16#2A;
   STAT5.STAT16[13] := B#16#29;
   STAT5.STAT16[14] := B#16#1;
   STAT5.STAT16[15] := B#16#0;
   STAT5.STAT16[16] := B#16#0;
   STAT5.STAT16[17] := B#16#0;
   STAT5.STAT16[18] := B#16#0;
   STAT5.STAT16[19] := B#16#0;
   STAT5.STAT16[20] := B#16#0;
   STAT5.STAT16[21] := B#16#0;
   STAT5.STAT16[22] := B#16#0;
   STAT5.STAT16[23] := B#16#0;
   STAT5.STAT16[24] := B#16#0;
   STAT5.STAT16[25] := B#16#0;
   STAT5.STAT16[26] := B#16#0;
   STAT5.STAT16[27] := B#16#0;
   STAT5.STAT16[28] := B#16#0;
   STAT5.STAT16[29] := B#16#0;
   STAT5.STAT16[30] := B#16#0;
   STAT5.STAT16[31] := B#16#0;
   STAT5.STAT16[32] := B#16#0;
   STAT5.STAT16[33] := B#16#0;
   STAT5.STAT16[34] := B#16#0;
   STAT5.STAT16[35] := B#16#0;
   STAT5.STAT16[36] := B#16#0;
   STAT5.STAT16[37] := B#16#0;
   STAT5.STAT16[38] := B#16#0;
   STAT5.STAT16[39] := B#16#0;
   STAT5.STAT16[40] := B#16#0;
   STAT5.STAT16[41] := B#16#0;
   STAT5.STAT16[42] := B#16#0;
   STAT5.STAT16[43] := B#16#0;
   STAT5.STAT16[44] := B#16#0;
   STAT5.STAT16[45] := B#16#0;
   STAT5.STAT16[46] := B#16#0;
   STAT5.STAT16[47] := B#16#0;
   STAT5.STAT16[48] := B#16#0;
   STAT5.STAT16[49] := B#16#0;
   STAT5.STAT16[50] := B#16#0;
   STAT5.STAT16[51] := B#16#0;
   STAT5.STAT16[52] := B#16#0;
   STAT5.STAT16[53] := B#16#0;
   STAT5.STAT16[54] := B#16#0;
   STAT5.STAT16[55] := B#16#0;
   STAT5.STAT16[56] := B#16#0;
   STAT5.STAT16[57] := B#16#0;
   STAT5.STAT16[58] := B#16#0;
   STAT5.STAT16[59] := B#16#0;
   STAT5.STAT16[60] := B#16#0;
   STAT5.STAT16[61] := B#16#0;
   STAT5.STAT16[62] := B#16#0;
   STAT5.STAT16[63] := B#16#0;
   STAT5.STAT16[64] := B#16#0;
   STAT5.STAT16[65] := B#16#0;
   STAT5.STAT16[66] := B#16#0;
   STAT5.STAT16[67] := B#16#0;
   STAT5.STAT16[68] := B#16#0;
   STAT5.STAT16[69] := B#16#0;
   STAT5.STAT16[70] := B#16#0;
   STAT5.STAT16[71] := B#16#0;
   STAT5.STAT16[72] := B#16#0;
   STAT5.STAT16[73] := B#16#0;
   STAT5.STAT16[74] := B#16#0;
   STAT5.STAT16[75] := B#16#0;
   STAT5.STAT16[76] := B#16#0;
   STAT5.STAT16[77] := B#16#0;
   STAT5.STAT16[78] := B#16#0;
   STAT5.STAT16[79] := B#16#0;
   STAT5.STAT16[80] := B#16#0;
   STAT5.STAT16[81] := B#16#0;
   STAT5.STAT16[82] := B#16#0;
   STAT5.STAT16[83] := B#16#0;
   STAT5.STAT16[84] := B#16#0;
   STAT5.STAT16[85] := B#16#0;
   STAT5.STAT16[86] := B#16#0;
   STAT5.STAT16[87] := B#16#0;
   STAT5.STAT16[88] := B#16#0;
   STAT5.STAT16[89] := B#16#0;
   STAT5.STAT16[90] := B#16#0;
   STAT5.STAT16[91] := B#16#0;
   STAT5.STAT16[92] := B#16#0;
   STAT5.STAT16[93] := B#16#0;
   STAT5.STAT16[94] := B#16#0;
   STAT5.STAT16[95] := B#16#0;
   STAT5.STAT16[96] := B#16#0;
   STAT5.STAT16[97] := B#16#0;
   STAT5.STAT16[98] := B#16#0;
   STAT5.STAT16[99] := B#16#0;
   STAT5.STAT16[100] := B#16#0;
   STAT5.STAT16[101] := B#16#0;
   STAT5.STAT16[102] := B#16#0;
   STAT5.STAT16[103] := B#16#0;
   STAT5.STAT16[104] := B#16#0;
   STAT5.STAT16[105] := B#16#0;
   STAT5.STAT16[106] := B#16#0;
   STAT5.STAT16[107] := B#16#0;
   STAT5.STAT16[108] := B#16#0;
   STAT5.STAT16[109] := B#16#0;
   STAT5.STAT16[110] := B#16#0;
   STAT5.STAT16[111] := B#16#0;
   STAT5.STAT16[112] := B#16#0;
   STAT5.STAT16[113] := B#16#0;
   STAT5.STAT16[114] := B#16#0;
   STAT5.STAT16[115] := B#16#0;
   STAT5.STAT16[116] := B#16#0;
   STAT5.STAT16[117] := B#16#0;
   STAT5.STAT16[118] := B#16#0;
   STAT5.STAT16[119] := B#16#0;
   STAT5.STAT16[120] := B#16#0;
   STAT5.STAT16[121] := B#16#0;
   STAT5.STAT16[122] := B#16#0;
   STAT5.STAT16[123] := B#16#0;
   STAT5.STAT16[124] := B#16#0;
   STAT5.STAT16[125] := B#16#0;
   STAT5.STAT16[126] := B#16#0;
   STAT5.STAT16[127] := B#16#0;
   STAT5.STAT16[128] := B#16#0;
   STAT5.STAT16[129] := B#16#0;
   STAT5.STAT16[130] := B#16#0;
   STAT5.STAT16[131] := B#16#0;
   STAT5.STAT16[132] := B#16#0;
   STAT5.STAT16[133] := B#16#0;
   STAT5.STAT16[134] := B#16#0;
   STAT5.STAT16[135] := B#16#0;
   STAT5.STAT16[136] := B#16#0;
   STAT5.STAT16[137] := B#16#0;
   STAT5.STAT16[138] := B#16#0;
   STAT5.STAT16[139] := B#16#0;
   STAT5.STAT16[140] := B#16#0;
   STAT5.STAT16[141] := B#16#0;
   STAT5.STAT16[142] := B#16#0;
   STAT5.STAT16[143] := B#16#0;
   STAT5.STAT16[144] := B#16#0;
   STAT5.STAT16[145] := B#16#0;
   STAT5.STAT16[146] := B#16#0;
   STAT5.STAT16[147] := B#16#0;
   STAT5.STAT16[148] := B#16#0;
   STAT5.STAT16[149] := B#16#0;
   STAT5.STAT16[150] := B#16#0;
   STAT5.STAT16[151] := B#16#0;
   STAT5.STAT16[152] := B#16#0;
   STAT5.STAT16[153] := B#16#0;
   STAT5.STAT16[154] := B#16#0;
   STAT5.STAT16[155] := B#16#0;
   STAT5.STAT16[156] := B#16#0;
   STAT5.STAT16[157] := B#16#0;
   STAT5.STAT16[158] := B#16#0;
   STAT5.STAT16[159] := B#16#0;
   STAT5.STAT16[160] := B#16#0;
   STAT5.STAT16[161] := B#16#0;
   STAT5.STAT16[162] := B#16#0;
   STAT5.STAT16[163] := B#16#0;
   STAT5.STAT16[164] := B#16#0;
   STAT5.STAT16[165] := B#16#0;
   STAT5.STAT16[166] := B#16#0;
   STAT5.STAT16[167] := B#16#0;
   STAT5.STAT16[168] := B#16#0;
   STAT5.STAT16[169] := B#16#0;
   STAT5.STAT16[170] := B#16#0;
   STAT5.STAT16[171] := B#16#0;
   STAT5.STAT16[172] := B#16#0;
   STAT5.STAT16[173] := B#16#0;
   STAT5.STAT16[174] := B#16#0;
   STAT5.STAT16[175] := B#16#0;
   STAT5.STAT16[176] := B#16#0;
   STAT5.STAT16[177] := B#16#0;
   STAT5.STAT16[178] := B#16#0;
   STAT5.STAT16[179] := B#16#0;
   STAT5.STAT16[180] := B#16#0;
   STAT5.STAT16[181] := B#16#0;
   STAT5.STAT16[182] := B#16#0;
   STAT5.STAT16[183] := B#16#0;
   STAT5.STAT16[184] := B#16#0;
   STAT5.STAT16[185] := B#16#0;
   STAT5.STAT16[186] := B#16#0;
   STAT5.STAT16[187] := B#16#0;
   STAT5.STAT16[188] := B#16#0;
   STAT5.STAT16[189] := B#16#0;
   STAT5.STAT16[190] := B#16#0;
   STAT5.STAT16[191] := B#16#0;
   STAT5.STAT16[192] := B#16#0;
   STAT5.STAT16[193] := B#16#0;
   STAT5.STAT16[194] := B#16#0;
   STAT5.STAT16[195] := B#16#0;
   STAT5.STAT16[196] := B#16#0;
   STAT5.STAT16[197] := B#16#0;
   STAT5.STAT16[198] := B#16#0;
   STAT5.STAT16[199] := B#16#0;
   STAT5.STAT16[200] := B#16#0;
   STAT5.STAT16[201] := B#16#0;
   STAT5.STAT16[202] := B#16#0;
   STAT5.STAT16[203] := B#16#0;
   STAT5.STAT16[204] := B#16#0;
   STAT5.STAT16[205] := B#16#0;
   STAT5.STAT16[206] := B#16#0;
   STAT5.STAT16[207] := B#16#0;
   STAT5.STAT16[208] := B#16#0;
   STAT5.STAT16[209] := B#16#0;
   STAT5.STAT16[210] := B#16#0;
   STAT5.STAT16[211] := B#16#0;
   STAT5.STAT16[212] := B#16#0;
   STAT5.STAT16[213] := B#16#0;
   STAT5.STAT16[214] := B#16#0;
   STAT5.STAT16[215] := B#16#0;
   STAT5.STAT16[216] := B#16#0;
   STAT5.STAT16[217] := B#16#0;
   STAT5.STAT16[218] := B#16#0;
   STAT5.STAT16[219] := B#16#0;
   STAT5.STAT16[220] := B#16#0;
   STAT5.STAT16[221] := B#16#0;
   STAT5.STAT16[222] := B#16#0;
   STAT5.STAT16[223] := B#16#0;
   STAT5.STAT16[224] := B#16#0;
   STAT5.STAT16[225] := B#16#0;
   STAT5.STAT16[226] := B#16#0;
   STAT5.STAT16[227] := B#16#0;
   STAT5.STAT16[228] := B#16#0;
   STAT5.STAT16[229] := B#16#0;
   STAT5.STAT16[230] := B#16#0;
END_DATA_BLOCK

DATA_BLOCK DB 104
VERSION : 0.1


  STRUCT
   STAT0 : BOOL ;
   STAT1 : BOOL ;
   STAT2 : BOOL ;
   STAT3 : WORD ;
   STAT4 : INT ;
   STAT5 : STRUCT
    STAT6 : BYTE ;
    STAT7 : BYTE ;
    STAT8 : BYTE ;
    STAT9 : BYTE ;
    STAT10 : BYTE ;
    STAT11 : BYTE ;
    STAT12 : BYTE ;
    STAT13 : BYTE ;
    STAT14 : BYTE ;
    STAT15 : BYTE ;
    STAT16 : ARRAY  [0 .. 230 ] OF BYTE ;
   END_STRUCT ;
  END_STRUCT ;
BEGIN
   STAT0 := TRUE;
   STAT1 := TRUE;
   STAT2 := FALSE;
   STAT3 := W#16#1FF5;
   STAT4 := 28673;
   STAT5.STAT6 := B#16#0;
   STAT5.STAT7 := B#16#C;
   STAT5.STAT8 := B#16#0;
   STAT5.STAT9 := B#16#2;
   STAT5.STAT10 := B#16#80;
   STAT5.STAT11 := B#16#1E;
   STAT5.STAT12 := B#16#43;
   STAT5.STAT13 := B#16#0;
   STAT5.STAT14 := B#16#0;
   STAT5.STAT15 := B#16#8;
   STAT5.STAT16[0] := B#16#82;
   STAT5.STAT16[1] := B#16#0;
   STAT5.STAT16[2] := B#16#0;
   STAT5.STAT16[3] := B#16#0;
   STAT5.STAT16[4] := B#16#0;
   STAT5.STAT16[5] := B#16#0;
   STAT5.STAT16[6] := B#16#0;
   STAT5.STAT16[7] := B#16#8;
   STAT5.STAT16[8] := B#16#9F;
   STAT5.STAT16[9] := B#16#0;
   STAT5.STAT16[10] := B#16#D0;
   STAT5.STAT16[11] := B#16#42;
   STAT5.STAT16[12] := B#16#2A;
   STAT5.STAT16[13] := B#16#29;
   STAT5.STAT16[14] := B#16#1;
   STAT5.STAT16[15] := B#16#0;
   STAT5.STAT16[16] := B#16#0;
   STAT5.STAT16[17] := B#16#0;
   STAT5.STAT16[18] := B#16#0;
   STAT5.STAT16[19] := B#16#0;
   STAT5.STAT16[20] := B#16#0;
   STAT5.STAT16[21] := B#16#0;
   STAT5.STAT16[22] := B#16#0;
   STAT5.STAT16[23] := B#16#0;
   STAT5.STAT16[24] := B#16#0;
   STAT5.STAT16[25] := B#16#0;
   STAT5.STAT16[26] := B#16#0;
   STAT5.STAT16[27] := B#16#0;
   STAT5.STAT16[28] := B#16#0;
   STAT5.STAT16[29] := B#16#0;
   STAT5.STAT16[30] := B#16#0;
   STAT5.STAT16[31] := B#16#0;
   STAT5.STAT16[32] := B#16#0;
   STAT5.STAT16[33] := B#16#0;
   STAT5.STAT16[34] := B#16#0;
   STAT5.STAT16[35] := B#16#0;
   STAT5.STAT16[36] := B#16#0;
   STAT5.STAT16[37] := B#16#0;
   STAT5.STAT16[38] := B#16#0;
   STAT5.STAT16[39] := B#16#0;
   STAT5.STAT16[40] := B#16#0;
   STAT5.STAT16[41] := B#16#0;
   STAT5.STAT16[42] := B#16#0;
   STAT5.STAT16[43] := B#16#0;
   STAT5.STAT16[44] := B#16#0;
   STAT5.STAT16[45] := B#16#0;
   STAT5.STAT16[46] := B#16#0;
   STAT5.STAT16[47] := B#16#0;
   STAT5.STAT16[48] := B#16#0;
   STAT5.STAT16[49] := B#16#0;
   STAT5.STAT16[50] := B#16#0;
   STAT5.STAT16[51] := B#16#0;
   STAT5.STAT16[52] := B#16#0;
   STAT5.STAT16[53] := B#16#0;
   STAT5.STAT16[54] := B#16#0;
   STAT5.STAT16[55] := B#16#0;
   STAT5.STAT16[56] := B#16#0;
   STAT5.STAT16[57] := B#16#0;
   STAT5.STAT16[58] := B#16#0;
   STAT5.STAT16[59] := B#16#0;
   STAT5.STAT16[60] := B#16#0;
   STAT5.STAT16[61] := B#16#0;
   STAT5.STAT16[62] := B#16#0;
   STAT5.STAT16[63] := B#16#0;
   STAT5.STAT16[64] := B#16#0;
   STAT5.STAT16[65] := B#16#0;
   STAT5.STAT16[66] := B#16#0;
   STAT5.STAT16[67] := B#16#0;
   STAT5.STAT16[68] := B#16#0;
   STAT5.STAT16[69] := B#16#0;
   STAT5.STAT16[70] := B#16#0;
   STAT5.STAT16[71] := B#16#0;
   STAT5.STAT16[72] := B#16#0;
   STAT5.STAT16[73] := B#16#0;
   STAT5.STAT16[74] := B#16#0;
   STAT5.STAT16[75] := B#16#0;
   STAT5.STAT16[76] := B#16#0;
   STAT5.STAT16[77] := B#16#0;
   STAT5.STAT16[78] := B#16#0;
   STAT5.STAT16[79] := B#16#0;
   STAT5.STAT16[80] := B#16#0;
   STAT5.STAT16[81] := B#16#0;
   STAT5.STAT16[82] := B#16#0;
   STAT5.STAT16[83] := B#16#0;
   STAT5.STAT16[84] := B#16#0;
   STAT5.STAT16[85] := B#16#0;
   STAT5.STAT16[86] := B#16#0;
   STAT5.STAT16[87] := B#16#0;
   STAT5.STAT16[88] := B#16#0;
   STAT5.STAT16[89] := B#16#0;
   STAT5.STAT16[90] := B#16#0;
   STAT5.STAT16[91] := B#16#0;
   STAT5.STAT16[92] := B#16#0;
   STAT5.STAT16[93] := B#16#0;
   STAT5.STAT16[94] := B#16#0;
   STAT5.STAT16[95] := B#16#0;
   STAT5.STAT16[96] := B#16#0;
   STAT5.STAT16[97] := B#16#0;
   STAT5.STAT16[98] := B#16#0;
   STAT5.STAT16[99] := B#16#0;
   STAT5.STAT16[100] := B#16#0;
   STAT5.STAT16[101] := B#16#0;
   STAT5.STAT16[102] := B#16#0;
   STAT5.STAT16[103] := B#16#0;
   STAT5.STAT16[104] := B#16#0;
   STAT5.STAT16[105] := B#16#0;
   STAT5.STAT16[106] := B#16#0;
   STAT5.STAT16[107] := B#16#0;
   STAT5.STAT16[108] := B#16#0;
   STAT5.STAT16[109] := B#16#0;
   STAT5.STAT16[110] := B#16#0;
   STAT5.STAT16[111] := B#16#0;
   STAT5.STAT16[112] := B#16#0;
   STAT5.STAT16[113] := B#16#0;
   STAT5.STAT16[114] := B#16#0;
   STAT5.STAT16[115] := B#16#0;
   STAT5.STAT16[116] := B#16#0;
   STAT5.STAT16[117] := B#16#0;
   STAT5.STAT16[118] := B#16#0;
   STAT5.STAT16[119] := B#16#0;
   STAT5.STAT16[120] := B#16#0;
   STAT5.STAT16[121] := B#16#0;
   STAT5.STAT16[122] := B#16#0;
   STAT5.STAT16[123] := B#16#0;
   STAT5.STAT16[124] := B#16#0;
   STAT5.STAT16[125] := B#16#0;
   STAT5.STAT16[126] := B#16#0;
   STAT5.STAT16[127] := B#16#0;
   STAT5.STAT16[128] := B#16#0;
   STAT5.STAT16[129] := B#16#0;
   STAT5.STAT16[130] := B#16#0;
   STAT5.STAT16[131] := B#16#0;
   STAT5.STAT16[132] := B#16#0;
   STAT5.STAT16[133] := B#16#0;
   STAT5.STAT16[134] := B#16#0;
   STAT5.STAT16[135] := B#16#0;
   STAT5.STAT16[136] := B#16#0;
   STAT5.STAT16[137] := B#16#0;
   STAT5.STAT16[138] := B#16#0;
   STAT5.STAT16[139] := B#16#0;
   STAT5.STAT16[140] := B#16#0;
   STAT5.STAT16[141] := B#16#0;
   STAT5.STAT16[142] := B#16#0;
   STAT5.STAT16[143] := B#16#0;
   STAT5.STAT16[144] := B#16#0;
   STAT5.STAT16[145] := B#16#0;
   STAT5.STAT16[146] := B#16#0;
   STAT5.STAT16[147] := B#16#0;
   STAT5.STAT16[148] := B#16#0;
   STAT5.STAT16[149] := B#16#0;
   STAT5.STAT16[150] := B#16#0;
   STAT5.STAT16[151] := B#16#0;
   STAT5.STAT16[152] := B#16#0;
   STAT5.STAT16[153] := B#16#0;
   STAT5.STAT16[154] := B#16#0;
   STAT5.STAT16[155] := B#16#0;
   STAT5.STAT16[156] := B#16#0;
   STAT5.STAT16[157] := B#16#0;
   STAT5.STAT16[158] := B#16#0;
   STAT5.STAT16[159] := B#16#0;
   STAT5.STAT16[160] := B#16#0;
   STAT5.STAT16[161] := B#16#0;
   STAT5.STAT16[162] := B#16#0;
   STAT5.STAT16[163] := B#16#0;
   STAT5.STAT16[164] := B#16#0;
   STAT5.STAT16[165] := B#16#0;
   STAT5.STAT16[166] := B#16#0;
   STAT5.STAT16[167] := B#16#0;
   STAT5.STAT16[168] := B#16#0;
   STAT5.STAT16[169] := B#16#0;
   STAT5.STAT16[170] := B#16#0;
   STAT5.STAT16[171] := B#16#0;
   STAT5.STAT16[172] := B#16#0;
   STAT5.STAT16[173] := B#16#0;
   STAT5.STAT16[174] := B#16#0;
   STAT5.STAT16[175] := B#16#0;
   STAT5.STAT16[176] := B#16#0;
   STAT5.STAT16[177] := B#16#0;
   STAT5.STAT16[178] := B#16#0;
   STAT5.STAT16[179] := B#16#0;
   STAT5.STAT16[180] := B#16#0;
   STAT5.STAT16[181] := B#16#0;
   STAT5.STAT16[182] := B#16#0;
   STAT5.STAT16[183] := B#16#0;
   STAT5.STAT16[184] := B#16#0;
   STAT5.STAT16[185] := B#16#0;
   STAT5.STAT16[186] := B#16#0;
   STAT5.STAT16[187] := B#16#0;
   STAT5.STAT16[188] := B#16#0;
   STAT5.STAT16[189] := B#16#0;
   STAT5.STAT16[190] := B#16#0;
   STAT5.STAT16[191] := B#16#0;
   STAT5.STAT16[192] := B#16#0;
   STAT5.STAT16[193] := B#16#0;
   STAT5.STAT16[194] := B#16#0;
   STAT5.STAT16[195] := B#16#0;
   STAT5.STAT16[196] := B#16#0;
   STAT5.STAT16[197] := B#16#0;
   STAT5.STAT16[198] := B#16#0;
   STAT5.STAT16[199] := B#16#0;
   STAT5.STAT16[200] := B#16#0;
   STAT5.STAT16[201] := B#16#0;
   STAT5.STAT16[202] := B#16#0;
   STAT5.STAT16[203] := B#16#0;
   STAT5.STAT16[204] := B#16#0;
   STAT5.STAT16[205] := B#16#0;
   STAT5.STAT16[206] := B#16#0;
   STAT5.STAT16[207] := B#16#0;
   STAT5.STAT16[208] := B#16#0;
   STAT5.STAT16[209] := B#16#0;
   STAT5.STAT16[210] := B#16#0;
   STAT5.STAT16[211] := B#16#0;
   STAT5.STAT16[212] := B#16#0;
   STAT5.STAT16[213] := B#16#0;
   STAT5.STAT16[214] := B#16#0;
   STAT5.STAT16[215] := B#16#0;
   STAT5.STAT16[216] := B#16#0;
   STAT5.STAT16[217] := B#16#0;
   STAT5.STAT16[218] := B#16#0;
   STAT5.STAT16[219] := B#16#0;
   STAT5.STAT16[220] := B#16#0;
   STAT5.STAT16[221] := B#16#0;
   STAT5.STAT16[222] := B#16#0;
   STAT5.STAT16[223] := B#16#0;
   STAT5.STAT16[224] := B#16#0;
   STAT5.STAT16[225] := B#16#0;
   STAT5.STAT16[226] := B#16#0;
   STAT5.STAT16[227] := B#16#0;
   STAT5.STAT16[228] := B#16#0;
   STAT5.STAT16[229] := B#16#0;
   STAT5.STAT16[230] := B#16#0;
END_DATA_BLOCK

DATA_BLOCK DB 106
VERSION : 0.1


  STRUCT
   STAT0 : BOOL ;
   STAT1 : BOOL ;
   STAT2 : BOOL ;
   STAT3 : WORD ;
   STAT4 : INT ;
   STAT5 : STRUCT
    STAT6 : BYTE ;
    STAT7 : BYTE ;
    STAT8 : BYTE ;
    STAT9 : BYTE ;
    STAT10 : BYTE ;
    STAT11 : BYTE ;
    STAT12 : BYTE ;
    STAT13 : BYTE ;
    STAT14 : BYTE ;
    STAT15 : BYTE ;
    STAT16 : ARRAY  [0 .. 230 ] OF BYTE ;
   END_STRUCT ;
  END_STRUCT ;
BEGIN
   STAT0 := TRUE;
   STAT1 := TRUE;
   STAT2 := TRUE;
   STAT3 := W#16#1FF3;
   STAT4 := 28674;
   STAT5.STAT6 := B#16#8;
   STAT5.STAT7 := B#16#C;
   STAT5.STAT8 := B#16#0;
   STAT5.STAT9 := B#16#2;
   STAT5.STAT10 := B#16#80;
   STAT5.STAT11 := B#16#52;
   STAT5.STAT12 := B#16#5F;
   STAT5.STAT13 := B#16#10;
   STAT5.STAT14 := B#16#0;
   STAT5.STAT15 := B#16#0;
   STAT5.STAT16[0] := B#16#0;
   STAT5.STAT16[1] := B#16#0;
   STAT5.STAT16[2] := B#16#0;
   STAT5.STAT16[3] := B#16#0;
   STAT5.STAT16[4] := B#16#0;
   STAT5.STAT16[5] := B#16#0;
   STAT5.STAT16[6] := B#16#0;
   STAT5.STAT16[7] := B#16#0;
   STAT5.STAT16[8] := B#16#0;
   STAT5.STAT16[9] := B#16#0;
   STAT5.STAT16[10] := B#16#0;
   STAT5.STAT16[11] := B#16#0;
   STAT5.STAT16[12] := B#16#0;
   STAT5.STAT16[13] := B#16#0;
   STAT5.STAT16[14] := B#16#0;
   STAT5.STAT16[15] := B#16#0;
   STAT5.STAT16[16] := B#16#0;
   STAT5.STAT16[17] := B#16#0;
   STAT5.STAT16[18] := B#16#0;
   STAT5.STAT16[19] := B#16#0;
   STAT5.STAT16[20] := B#16#0;
   STAT5.STAT16[21] := B#16#0;
   STAT5.STAT16[22] := B#16#0;
   STAT5.STAT16[23] := B#16#0;
   STAT5.STAT16[24] := B#16#0;
   STAT5.STAT16[25] := B#16#0;
   STAT5.STAT16[26] := B#16#0;
   STAT5.STAT16[27] := B#16#3F;
   STAT5.STAT16[28] := B#16#82;
   STAT5.STAT16[29] := B#16#0;
   STAT5.STAT16[30] := B#16#0;
   STAT5.STAT16[31] := B#16#0;
   STAT5.STAT16[32] := B#16#1;
   STAT5.STAT16[33] := B#16#0;
   STAT5.STAT16[34] := B#16#0;
   STAT5.STAT16[35] := B#16#0;
   STAT5.STAT16[36] := B#16#0;
   STAT5.STAT16[37] := B#16#0;
   STAT5.STAT16[38] := B#16#0;
   STAT5.STAT16[39] := B#16#0;
   STAT5.STAT16[40] := B#16#0;
   STAT5.STAT16[41] := B#16#0;
   STAT5.STAT16[42] := B#16#0;
   STAT5.STAT16[43] := B#16#0;
   STAT5.STAT16[44] := B#16#0;
   STAT5.STAT16[45] := B#16#0;
   STAT5.STAT16[46] := B#16#0;
   STAT5.STAT16[47] := B#16#0;
   STAT5.STAT16[48] := B#16#0;
   STAT5.STAT16[49] := B#16#0;
   STAT5.STAT16[50] := B#16#0;
   STAT5.STAT16[51] := B#16#0;
   STAT5.STAT16[52] := B#16#0;
   STAT5.STAT16[53] := B#16#0;
   STAT5.STAT16[54] := B#16#0;
   STAT5.STAT16[55] := B#16#0;
   STAT5.STAT16[56] := B#16#0;
   STAT5.STAT16[57] := B#16#0;
   STAT5.STAT16[58] := B#16#0;
   STAT5.STAT16[59] := B#16#0;
   STAT5.STAT16[60] := B#16#0;
   STAT5.STAT16[61] := B#16#0;
   STAT5.STAT16[62] := B#16#0;
   STAT5.STAT16[63] := B#16#0;
   STAT5.STAT16[64] := B#16#0;
   STAT5.STAT16[65] := B#16#0;
   STAT5.STAT16[66] := B#16#0;
   STAT5.STAT16[67] := B#16#0;
   STAT5.STAT16[68] := B#16#0;
   STAT5.STAT16[69] := B#16#0;
   STAT5.STAT16[70] := B#16#0;
   STAT5.STAT16[71] := B#16#0;
   STAT5.STAT16[72] := B#16#0;
   STAT5.STAT16[73] := B#16#0;
   STAT5.STAT16[74] := B#16#0;
   STAT5.STAT16[75] := B#16#0;
   STAT5.STAT16[76] := B#16#0;
   STAT5.STAT16[77] := B#16#0;
   STAT5.STAT16[78] := B#16#0;
   STAT5.STAT16[79] := B#16#0;
   STAT5.STAT16[80] := B#16#0;
   STAT5.STAT16[81] := B#16#0;
   STAT5.STAT16[82] := B#16#0;
   STAT5.STAT16[83] := B#16#0;
   STAT5.STAT16[84] := B#16#0;
   STAT5.STAT16[85] := B#16#0;
   STAT5.STAT16[86] := B#16#0;
   STAT5.STAT16[87] := B#16#0;
   STAT5.STAT16[88] := B#16#0;
   STAT5.STAT16[89] := B#16#0;
   STAT5.STAT16[90] := B#16#3C;
   STAT5.STAT16[91] := B#16#81;
   STAT5.STAT16[92] := B#16#0;
   STAT5.STAT16[93] := B#16#0;
   STAT5.STAT16[94] := B#16#0;
   STAT5.STAT16[95] := B#16#8;
   STAT5.STAT16[96] := B#16#0;
   STAT5.STAT16[97] := B#16#0;
   STAT5.STAT16[98] := B#16#0;
   STAT5.STAT16[99] := B#16#0;
   STAT5.STAT16[100] := B#16#0;
   STAT5.STAT16[101] := B#16#0;
   STAT5.STAT16[102] := B#16#0;
   STAT5.STAT16[103] := B#16#0;
   STAT5.STAT16[104] := B#16#0;
   STAT5.STAT16[105] := B#16#0;
   STAT5.STAT16[106] := B#16#0;
   STAT5.STAT16[107] := B#16#0;
   STAT5.STAT16[108] := B#16#0;
   STAT5.STAT16[109] := B#16#0;
   STAT5.STAT16[110] := B#16#0;
   STAT5.STAT16[111] := B#16#C;
   STAT5.STAT16[112] := B#16#0;
   STAT5.STAT16[113] := B#16#0;
   STAT5.STAT16[114] := B#16#0;
   STAT5.STAT16[115] := B#16#0;
   STAT5.STAT16[116] := B#16#0;
   STAT5.STAT16[117] := B#16#0;
   STAT5.STAT16[118] := B#16#0;
   STAT5.STAT16[119] := B#16#0;
   STAT5.STAT16[120] := B#16#0;
   STAT5.STAT16[121] := B#16#0;
   STAT5.STAT16[122] := B#16#0;
   STAT5.STAT16[123] := B#16#0;
   STAT5.STAT16[124] := B#16#0;
   STAT5.STAT16[125] := B#16#0;
   STAT5.STAT16[126] := B#16#C0;
   STAT5.STAT16[127] := B#16#82;
   STAT5.STAT16[128] := B#16#0;
   STAT5.STAT16[129] := B#16#0;
   STAT5.STAT16[130] := B#16#0;
   STAT5.STAT16[131] := B#16#0;
   STAT5.STAT16[132] := B#16#0;
   STAT5.STAT16[133] := B#16#2;
   STAT5.STAT16[134] := B#16#0;
   STAT5.STAT16[135] := B#16#0;
   STAT5.STAT16[136] := B#16#0;
   STAT5.STAT16[137] := B#16#0;
   STAT5.STAT16[138] := B#16#0;
   STAT5.STAT16[139] := B#16#0;
   STAT5.STAT16[140] := B#16#0;
   STAT5.STAT16[141] := B#16#0;
   STAT5.STAT16[142] := B#16#0;
   STAT5.STAT16[143] := B#16#0;
   STAT5.STAT16[144] := B#16#0;
   STAT5.STAT16[145] := B#16#0;
   STAT5.STAT16[146] := B#16#0;
   STAT5.STAT16[147] := B#16#0;
   STAT5.STAT16[148] := B#16#0;
   STAT5.STAT16[149] := B#16#0;
   STAT5.STAT16[150] := B#16#8;
   STAT5.STAT16[151] := B#16#9F;
   STAT5.STAT16[152] := B#16#0;
   STAT5.STAT16[153] := B#16#C8;
   STAT5.STAT16[154] := B#16#42;
   STAT5.STAT16[155] := B#16#2A;
   STAT5.STAT16[156] := B#16#29;
   STAT5.STAT16[157] := B#16#1;
   STAT5.STAT16[158] := B#16#12;
   STAT5.STAT16[159] := B#16#1;
   STAT5.STAT16[160] := B#16#3;
   STAT5.STAT16[161] := B#16#D1;
   STAT5.STAT16[162] := B#16#8;
   STAT5.STAT16[163] := B#16#C;
   STAT5.STAT16[164] := B#16#0;
   STAT5.STAT16[165] := B#16#7D;
   STAT5.STAT16[166] := B#16#81;
   STAT5.STAT16[167] := B#16#76;
   STAT5.STAT16[168] := B#16#42;
   STAT5.STAT16[169] := B#16#2;
   STAT5.STAT16[170] := B#16#6;
   STAT5.STAT16[171] := B#16#82;
   STAT5.STAT16[172] := B#16#0;
   STAT5.STAT16[173] := B#16#0;
   STAT5.STAT16[174] := B#16#4;
   STAT5.STAT16[175] := B#16#0;
   STAT5.STAT16[176] := B#16#0;
   STAT5.STAT16[177] := B#16#0;
   STAT5.STAT16[178] := B#16#0;
   STAT5.STAT16[179] := B#16#0;
   STAT5.STAT16[180] := B#16#0;
   STAT5.STAT16[181] := B#16#0;
   STAT5.STAT16[182] := B#16#0;
   STAT5.STAT16[183] := B#16#0;
   STAT5.STAT16[184] := B#16#0;
   STAT5.STAT16[185] := B#16#0;
   STAT5.STAT16[186] := B#16#0;
   STAT5.STAT16[187] := B#16#0;
   STAT5.STAT16[188] := B#16#0;
   STAT5.STAT16[189] := B#16#0;
   STAT5.STAT16[190] := B#16#0;
   STAT5.STAT16[191] := B#16#0;
   STAT5.STAT16[192] := B#16#0;
   STAT5.STAT16[193] := B#16#0;
   STAT5.STAT16[194] := B#16#0;
   STAT5.STAT16[195] := B#16#0;
   STAT5.STAT16[196] := B#16#0;
   STAT5.STAT16[197] := B#16#0;
   STAT5.STAT16[198] := B#16#0;
   STAT5.STAT16[199] := B#16#0;
   STAT5.STAT16[200] := B#16#0;
   STAT5.STAT16[201] := B#16#0;
   STAT5.STAT16[202] := B#16#0;
   STAT5.STAT16[203] := B#16#0;
   STAT5.STAT16[204] := B#16#0;
   STAT5.STAT16[205] := B#16#0;
   STAT5.STAT16[206] := B#16#0;
   STAT5.STAT16[207] := B#16#0;
   STAT5.STAT16[208] := B#16#0;
   STAT5.STAT16[209] := B#16#0;
   STAT5.STAT16[210] := B#16#0;
   STAT5.STAT16[211] := B#16#0;
   STAT5.STAT16[212] := B#16#0;
   STAT5.STAT16[213] := B#16#0;
   STAT5.STAT16[214] := B#16#0;
   STAT5.STAT16[215] := B#16#0;
   STAT5.STAT16[216] := B#16#0;
   STAT5.STAT16[217] := B#16#0;
   STAT5.STAT16[218] := B#16#0;
   STAT5.STAT16[219] := B#16#0;
   STAT5.STAT16[220] := B#16#0;
   STAT5.STAT16[221] := B#16#0;
   STAT5.STAT16[222] := B#16#0;
   STAT5.STAT16[223] := B#16#0;
   STAT5.STAT16[224] := B#16#0;
   STAT5.STAT16[225] := B#16#0;
   STAT5.STAT16[226] := B#16#0;
   STAT5.STAT16[227] := B#16#0;
   STAT5.STAT16[228] := B#16#0;
   STAT5.STAT16[229] := B#16#0;
   STAT5.STAT16[230] := B#16#0;
END_DATA_BLOCK

FUNCTION_BLOCK FB 500
VERSION : 0.1


VAR_INPUT
  IN0 : BOOL ;
  IN1 : BOOL ;
  IN2 : BOOL ;
END_VAR
VAR_OUTPUT
  OUT3 : BOOL ;
  OUT4 : BOOL ;
END_VAR
VAR
  STAT5 : BOOL ;
  STAT6 : BOOL ;
  STAT7 : BOOL ;
  STAT8 : BOOL ;
END_VAR
BEGIN
NETWORK
TITLE =
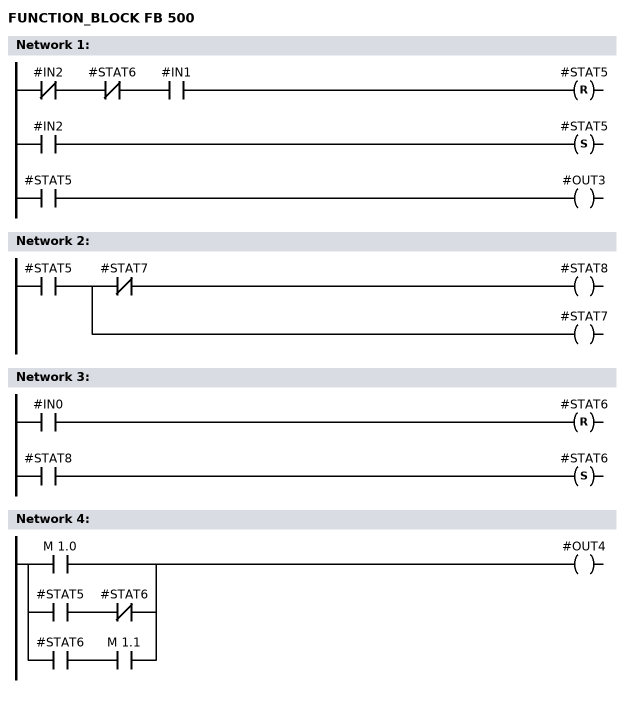

      AN    #IN2;
      AN    #STAT6;
      A     #IN1;
      R     #STAT5;
      A     #IN2;
      S     #STAT5;
      A     #STAT5;
      =     #OUT3;
NETWORK
TITLE =

      A     #STAT5;
      =     L      0.0;
      A     L      0.0;
      AN    #STAT7;
      =     #STAT8;
      A     L      0.0;
      BLD   102;
      =     #STAT7;
NETWORK
TITLE =

      A     #IN0;
      R     #STAT6;
      A     #STAT8;
      S     #STAT6;
      NOP   0;
NETWORK
TITLE =

      O     M      1.0;
      O     ;
      A     #STAT5;
      AN    #STAT6;
      O     ;
      A     #STAT6;
      A     M      1.1;
      =     #OUT4;
END_FUNCTION_BLOCK

FUNCTION FC 0 : VOID
VERSION : 0.1

BEGIN
NETWORK
TITLE =
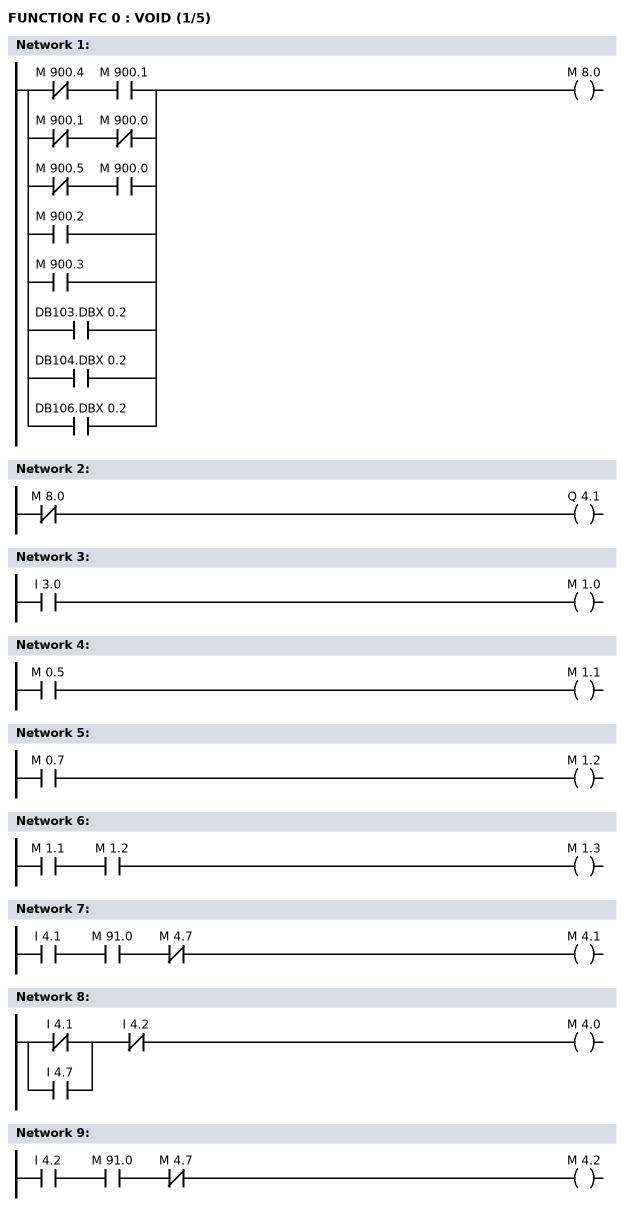

      AN    M    900.4;
      A     M    900.1;
      O     ;
      AN    M    900.1;
      AN    M    900.0;
      O     ;
      AN    M    900.5;
      A     M    900.0;
      O     M    900.2;
      O     M    900.3;
      O     DB103.DBX    0.2;
      O     DB104.DBX    0.2;
      O     DB106.DBX    0.2;
      =     M      8.0;
NETWORK
TITLE =

      AN    M      8.0;
      =     Q      4.1;
NETWORK
TITLE =

      A     I      3.0;
      =     M      1.0;
NETWORK
TITLE =

      A     M      0.5;
      =     M      1.1;
NETWORK
TITLE =

      A     M      0.7;
      =     M      1.2;
NETWORK
TITLE =

      A     M      1.1;
      A     M      1.2;
      =     M      1.3;
NETWORK
TITLE =

      A     I      4.1;
      A     M     91.0;
      AN    M      4.7;
      =     M      4.1;
NETWORK
TITLE =

      A(    ;
      ON    I      4.1;
      O     I      4.7;
      )     ;
      AN    I      4.2;
      =     M      4.0;
NETWORK
TITLE =

      A     I      4.2;
      A     M     91.0;
      AN    M      4.7;
      =     M      4.2;
NETWORK
TITLE =
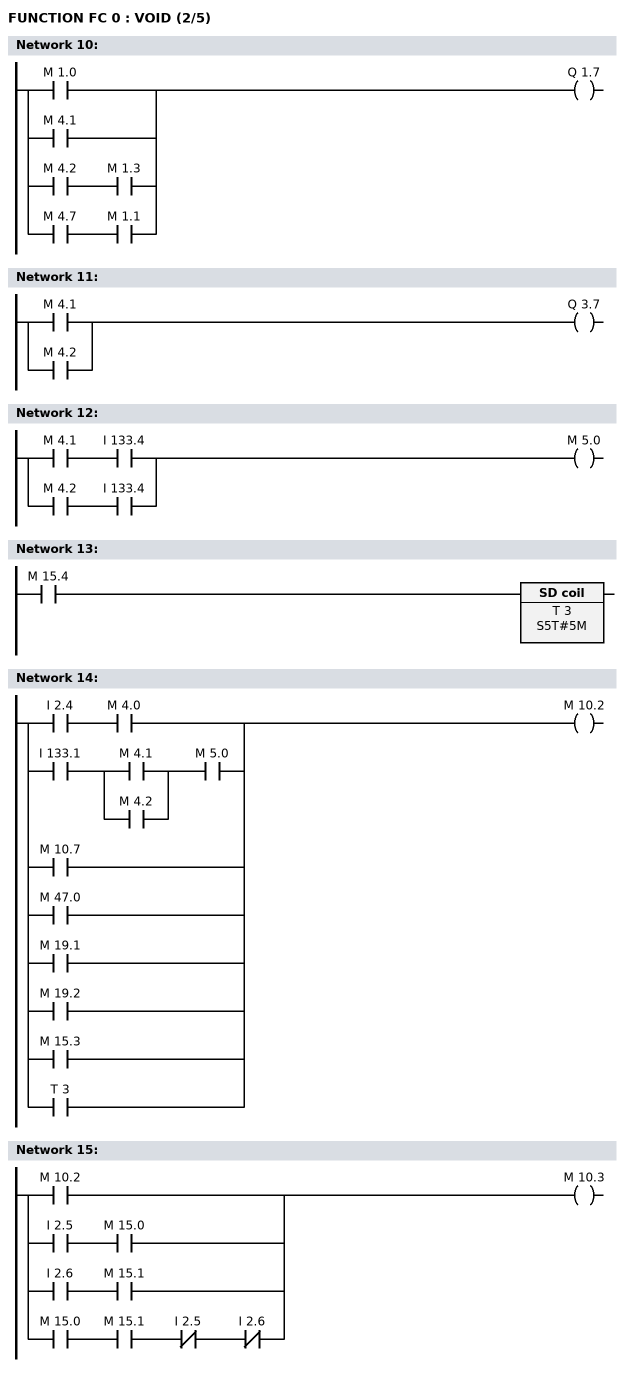

      O     M      1.0;
      O     M      4.1;
      O     ;
      A     M      4.2;
      A     M      1.3;
      O     ;
      A     M      4.7;
      A     M      1.1;
      =     Q      1.7;
NETWORK
TITLE =

      O     M      4.1;
      O     M      4.2;
      =     Q      3.7;
NETWORK
TITLE =

      A     M      4.1;
      A     I    133.4;
      O     ;
      A     M      4.2;
      A     I    133.4;
      =     M      5.0;
NETWORK
TITLE =

      A     M     15.4;
      L     S5T#5M;
      SD    T      3;
      NOP   0;
      NOP   0;
      NOP   0;
      NOP   0;
NETWORK
TITLE =

      A     I      2.4;
      A     M      4.0;
      O     ;
      A     I    133.1;
      A(    ;
      O     M      4.1;
      O     M      4.2;
      )     ;
      A     M      5.0;
      O     M     10.7;
      O     M     47.0;
      O     M     19.1;
      O     M     19.2;
      O     M     15.3;
      O     T      3;
      =     M     10.2;
NETWORK
TITLE =

      O     M     10.2;
      O     ;
      A     I      2.5;
      A     M     15.0;
      O     ;
      A     I      2.6;
      A     M     15.1;
      O     ;
      A     M     15.0;
      A     M     15.1;
      AN    I      2.5;
      AN    I      2.6;
      =     M     10.3;
NETWORK
TITLE =
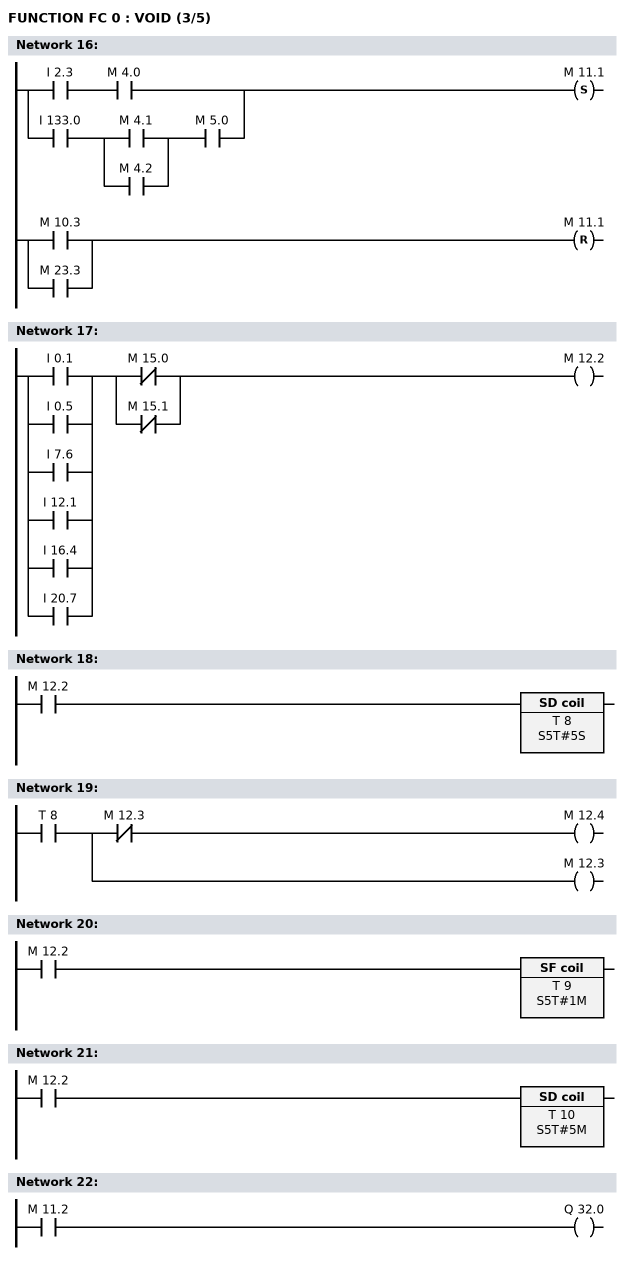

      A(    ;
      A     I      2.3;
      A     M      4.0;
      O     ;
      A     I    133.0;
      A(    ;
      O     M      4.1;
      O     M      4.2;
      )     ;
      A     M      5.0;
      )     ;
      S     M     11.1;
      A(    ;
      O     M     10.3;
      O     M     23.3;
      )     ;
      R     M     11.1;
      NOP   0;
NETWORK
TITLE =

      A(    ;
      O     I      0.1;
      O     I      0.5;
      O     I      7.6;
      O     I     12.1;
      O     I     16.4;
      O     I     20.7;
      )     ;
      A(    ;
      ON    M     15.0;
      ON    M     15.1;
      )     ;
      =     M     12.2;
NETWORK
TITLE =

      A     M     12.2;
      L     S5T#5S;
      SD    T      8;
      NOP   0;
      NOP   0;
      NOP   0;
      NOP   0;
NETWORK
TITLE =

      A     T      8;
      =     L      0.0;
      A     L      0.0;
      AN    M     12.3;
      =     M     12.4;
      A     L      0.0;
      BLD   102;
      =     M     12.3;
NETWORK
TITLE =

      A     M     12.2;
      L     S5T#1M;
      SF    T      9;
      NOP   0;
      NOP   0;
      NOP   0;
      NOP   0;
NETWORK
TITLE =

      A     M     12.2;
      L     S5T#5M;
      SD    T     10;
      NOP   0;
      NOP   0;
      NOP   0;
      NOP   0;
NETWORK
TITLE =

      A     M     11.2;
      =     Q     32.0;
NETWORK
TITLE =
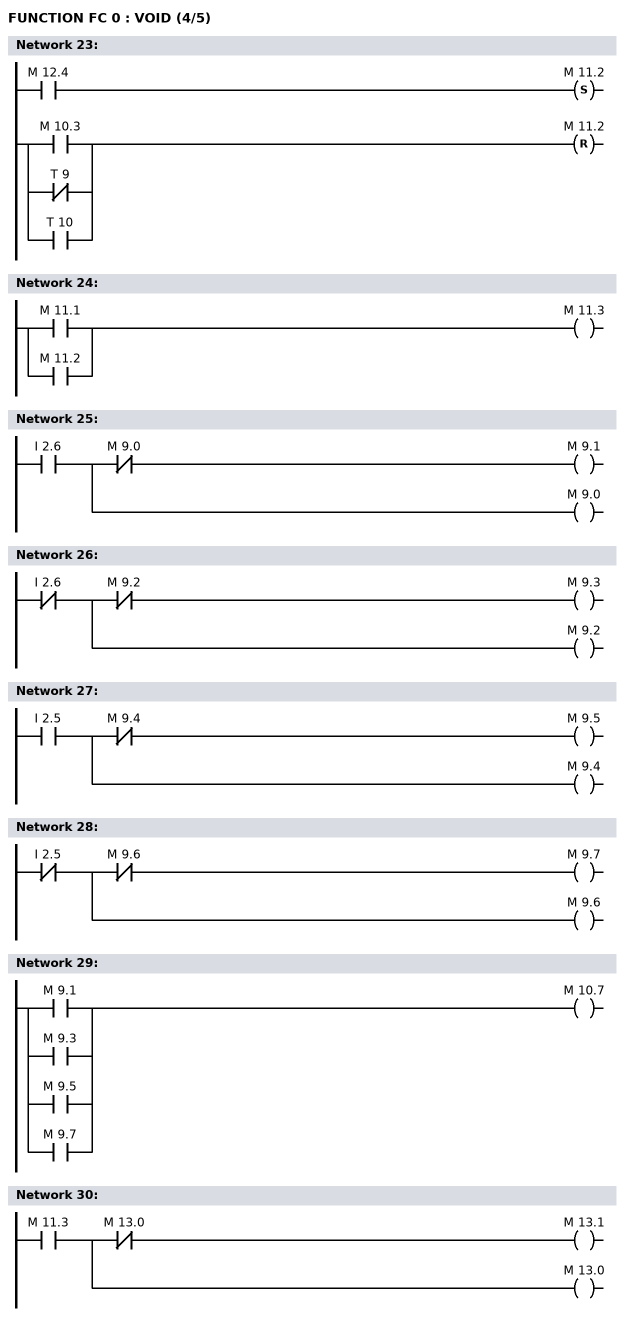

      A     M     12.4;
      S     M     11.2;
      A(    ;
      O     M     10.3;
      ON    T      9;
      O     T     10;
      )     ;
      R     M     11.2;
      NOP   0;
NETWORK
TITLE =

      O     M     11.1;
      O     M     11.2;
      =     M     11.3;
NETWORK
TITLE =

      A     I      2.6;
      =     L      0.0;
      A     L      0.0;
      AN    M      9.0;
      =     M      9.1;
      A     L      0.0;
      BLD   102;
      =     M      9.0;
NETWORK
TITLE =

      AN    I      2.6;
      =     L      0.0;
      A     L      0.0;
      AN    M      9.2;
      =     M      9.3;
      A     L      0.0;
      BLD   102;
      =     M      9.2;
NETWORK
TITLE =

      A     I      2.5;
      =     L      0.0;
      A     L      0.0;
      AN    M      9.4;
      =     M      9.5;
      A     L      0.0;
      BLD   102;
      =     M      9.4;
NETWORK
TITLE =

      AN    I      2.5;
      =     L      0.0;
      A     L      0.0;
      AN    M      9.6;
      =     M      9.7;
      A     L      0.0;
      BLD   102;
      =     M      9.6;
NETWORK
TITLE =

      O     M      9.1;
      O     M      9.3;
      O     M      9.5;
      O     M      9.7;
      =     M     10.7;
NETWORK
TITLE =

      A     M     11.3;
      =     L      0.0;
      A     L      0.0;
      AN    M     13.0;
      =     M     13.1;
      A     L      0.0;
      BLD   102;
      =     M     13.0;
NETWORK
TITLE =
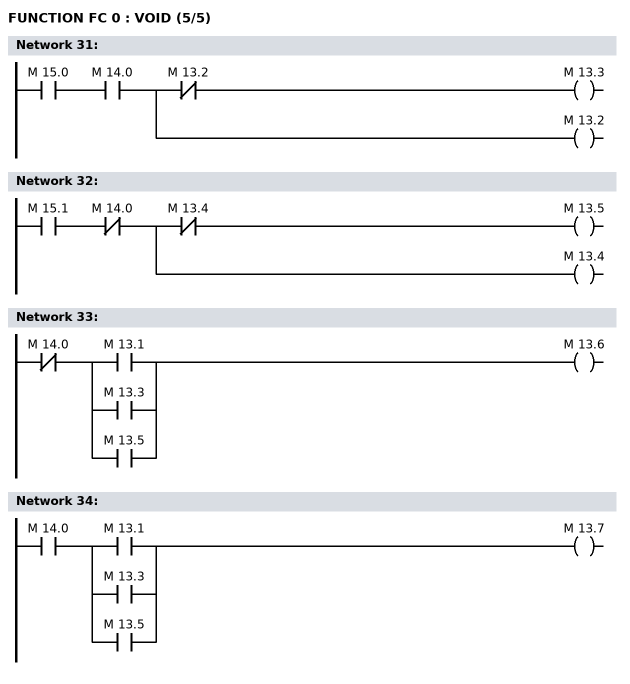

      A     M     15.0;
      A     M     14.0;
      =     L      0.0;
      A     L      0.0;
      AN    M     13.2;
      =     M     13.3;
      A     L      0.0;
      BLD   102;
      =     M     13.2;
NETWORK
TITLE =

      A     M     15.1;
      AN    M     14.0;
      =     L      0.0;
      A     L      0.0;
      AN    M     13.4;
      =     M     13.5;
      A     L      0.0;
      BLD   102;
      =     M     13.4;
NETWORK
TITLE =

      AN    M     14.0;
      A(    ;
      O     M     13.1;
      O     M     13.3;
      O     M     13.5;
      )     ;
      =     M     13.6;
NETWORK
TITLE =

      A     M     14.0;
      A(    ;
      O     M     13.1;
      O     M     13.3;
      O     M     13.5;
      )     ;
      =     M     13.7;
NETWORK
TITLE =

      A(    ;
      A     M     13.7;
      R     M     14.0;
      A     M     13.6;
      S     M     14.0;
      A     M     14.0;
      )     ;
      AN    I      2.5;
      AN    I      2.6;
      O     I      2.5;
      =     M     14.2;
NETWORK
TITLE =
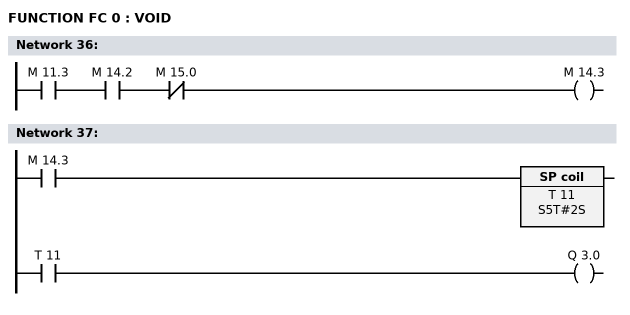

      A     M     11.3;
      A     M     14.2;
      AN    M     15.0;
      =     M     14.3;
NETWORK
TITLE =

      A     M     14.3;
      L     S5T#2S;
      SP    T     11;
      NOP   0;
      NOP   0;
      NOP   0;
      A     T     11;
      =     Q      3.0;
NETWORK
TITLE =

      A(    ;
      AN    M     14.3;
      L     S5T#2S;
      SP    T     12;
      NOP   0;
      NOP   0;
      NOP   0;
      A     T     12;
      )     ;
      NOT   ;
      AN    M     19.1;
      AN    M     19.2;
      AN    M     15.3;
      =     Q      3.1;
NETWORK
TITLE =
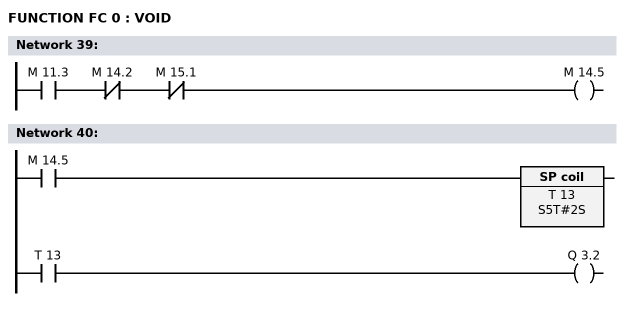

      A     M     11.3;
      AN    M     14.2;
      AN    M     15.1;
      =     M     14.5;
NETWORK
TITLE =

      A     M     14.5;
      L     S5T#2S;
      SP    T     13;
      NOP   0;
      NOP   0;
      NOP   0;
      A     T     13;
      =     Q      3.2;
NETWORK
TITLE =

      A(    ;
      AN    M     14.5;
      L     S5T#2S;
      SP    T     14;
      NOP   0;
      NOP   0;
      NOP   0;
      A     T     14;
      )     ;
      NOT   ;
      AN    M     19.1;
      AN    M     19.2;
      AN    M     15.3;
      =     Q      3.3;
NETWORK
TITLE =
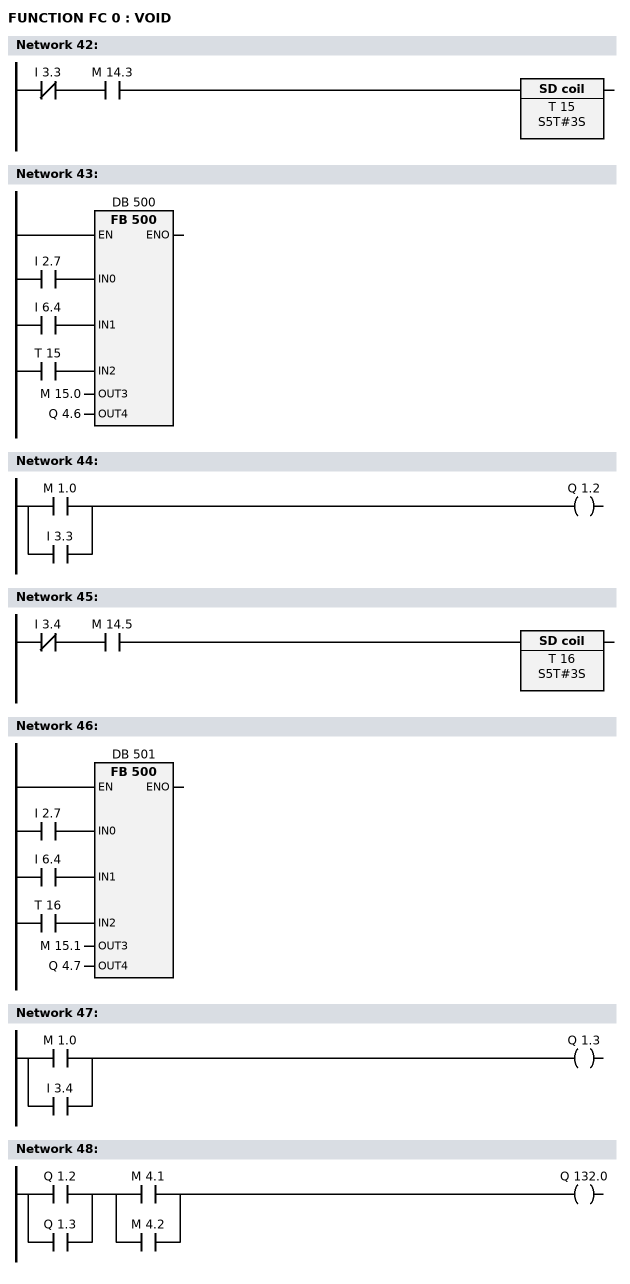

      AN    I      3.3;
      A     M     14.3;
      L     S5T#3S;
      SD    T     15;
      NOP   0;
      NOP   0;
      NOP   0;
      NOP   0;
NETWORK
TITLE =

      A     I      2.7;
      =     L      0.0;
      BLD   103;
      A     I      6.4;
      =     L      0.1;
      BLD   103;
      A     T     15;
      =     L      0.2;
      BLD   103;
      CALL FB   500 , DB   500 (
           IN0                      := L      0.0,
           IN1                      := L      0.1,
           IN2                      := L      0.2,
           OUT3                     := M     15.0,
           OUT4                     := Q      4.6);
      NOP   0;
NETWORK
TITLE =

      O     M      1.0;
      O     I      3.3;
      =     Q      1.2;
NETWORK
TITLE =

      AN    I      3.4;
      A     M     14.5;
      L     S5T#3S;
      SD    T     16;
      NOP   0;
      NOP   0;
      NOP   0;
      NOP   0;
NETWORK
TITLE =

      A     I      2.7;
      =     L      0.0;
      BLD   103;
      A     I      6.4;
      =     L      0.1;
      BLD   103;
      A     T     16;
      =     L      0.2;
      BLD   103;
      CALL FB   500 , DB   501 (
           IN0                      := L      0.0,
           IN1                      := L      0.1,
           IN2                      := L      0.2,
           OUT3                     := M     15.1,
           OUT4                     := Q      4.7);
      NOP   0;
NETWORK
TITLE =

      O     M      1.0;
      O     I      3.4;
      =     Q      1.3;
NETWORK
TITLE =

      A(    ;
      O     Q      1.2;
      O     Q      1.3;
      )     ;
      A(    ;
      O     M      4.1;
      O     M      4.2;
      )     ;
      =     Q    132.0;
NETWORK
TITLE =

      A(    ;
      AN    I      0.2;
      L     S5T#2S;
      SD    T     17;
      NOP   0;
      NOP   0;
      NOP   0;
      A     T     17;
      )     ;
      NOT   ;
      =     Q      2.4;
NETWORK
TITLE =
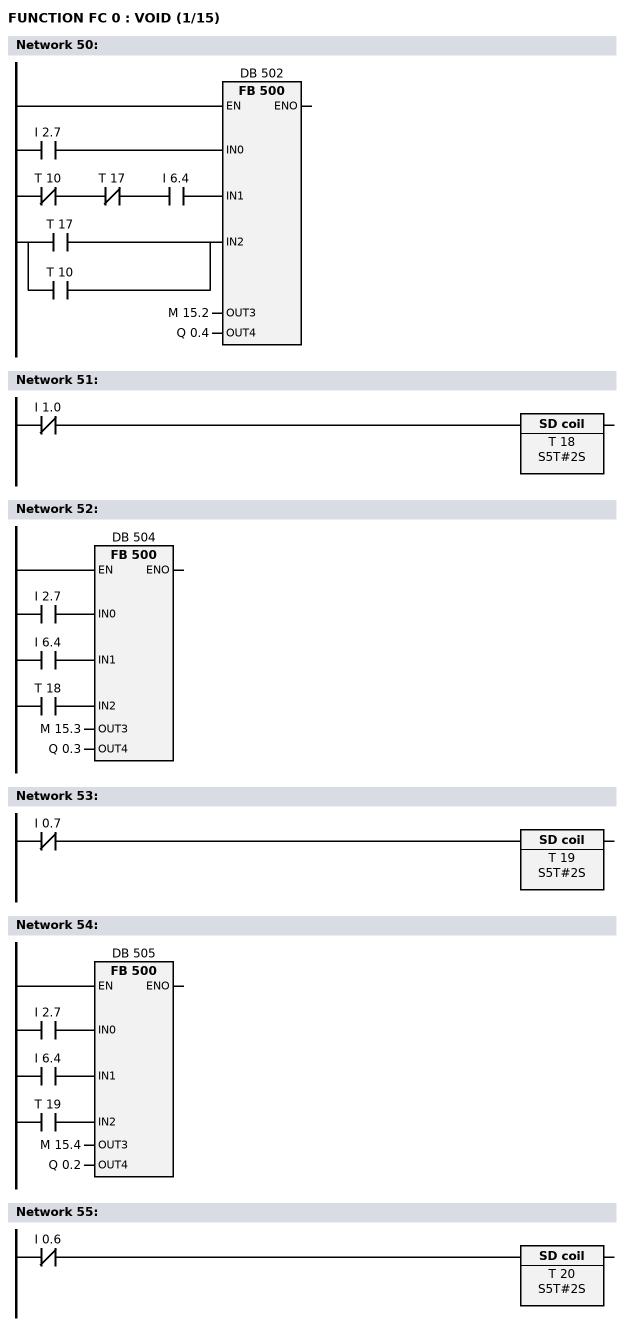

      A     I      2.7;
      =     L      0.0;
      BLD   103;
      AN    T     10;
      AN    T     17;
      A     I      6.4;
      =     L      0.1;
      BLD   103;
      A(    ;
      O     T     17;
      O     T     10;
      )     ;
      =     L      0.2;
      BLD   103;
      CALL FB   500 , DB   502 (
           IN0                      := L      0.0,
           IN1                      := L      0.1,
           IN2                      := L      0.2,
           OUT3                     := M     15.2,
           OUT4                     := Q      0.4);
      NOP   0;
NETWORK
TITLE =

      AN    I      1.0;
      L     S5T#2S;
      SD    T     18;
      NOP   0;
      NOP   0;
      NOP   0;
      NOP   0;
NETWORK
TITLE =

      A     I      2.7;
      =     L      0.0;
      BLD   103;
      A     I      6.4;
      =     L      0.1;
      BLD   103;
      A     T     18;
      =     L      0.2;
      BLD   103;
      CALL FB   500 , DB   504 (
           IN0                      := L      0.0,
           IN1                      := L      0.1,
           IN2                      := L      0.2,
           OUT3                     := M     15.3,
           OUT4                     := Q      0.3);
      NOP   0;
NETWORK
TITLE =

      AN    I      0.7;
      L     S5T#2S;
      SD    T     19;
      NOP   0;
      NOP   0;
      NOP   0;
      NOP   0;
NETWORK
TITLE =

      A     I      2.7;
      =     L      0.0;
      BLD   103;
      A     I      6.4;
      =     L      0.1;
      BLD   103;
      A     T     19;
      =     L      0.2;
      BLD   103;
      CALL FB   500 , DB   505 (
           IN0                      := L      0.0,
           IN1                      := L      0.1,
           IN2                      := L      0.2,
           OUT3                     := M     15.4,
           OUT4                     := Q      0.2);
      NOP   0;
NETWORK
TITLE =

      AN    I      0.6;
      L     S5T#2S;
      SD    T     20;
      NOP   0;
      NOP   0;
      NOP   0;
      NOP   0;
NETWORK
TITLE =
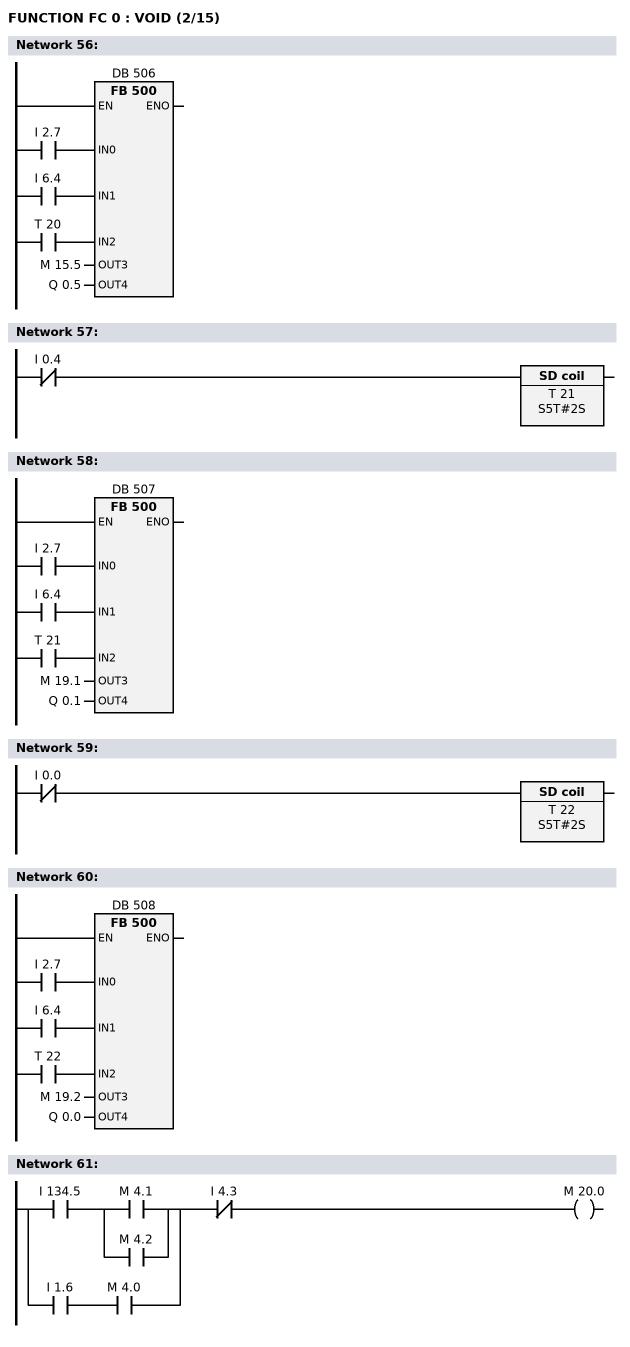

      A     I      2.7;
      =     L      0.0;
      BLD   103;
      A     I      6.4;
      =     L      0.1;
      BLD   103;
      A     T     20;
      =     L      0.2;
      BLD   103;
      CALL FB   500 , DB   506 (
           IN0                      := L      0.0,
           IN1                      := L      0.1,
           IN2                      := L      0.2,
           OUT3                     := M     15.5,
           OUT4                     := Q      0.5);
      NOP   0;
NETWORK
TITLE =

      AN    I      0.4;
      L     S5T#2S;
      SD    T     21;
      NOP   0;
      NOP   0;
      NOP   0;
      NOP   0;
NETWORK
TITLE =

      A     I      2.7;
      =     L      0.0;
      BLD   103;
      A     I      6.4;
      =     L      0.1;
      BLD   103;
      A     T     21;
      =     L      0.2;
      BLD   103;
      CALL FB   500 , DB   507 (
           IN0                      := L      0.0,
           IN1                      := L      0.1,
           IN2                      := L      0.2,
           OUT3                     := M     19.1,
           OUT4                     := Q      0.1);
      NOP   0;
NETWORK
TITLE =

      AN    I      0.0;
      L     S5T#2S;
      SD    T     22;
      NOP   0;
      NOP   0;
      NOP   0;
      NOP   0;
NETWORK
TITLE =

      A     I      2.7;
      =     L      0.0;
      BLD   103;
      A     I      6.4;
      =     L      0.1;
      BLD   103;
      A     T     22;
      =     L      0.2;
      BLD   103;
      CALL FB   500 , DB   508 (
           IN0                      := L      0.0,
           IN1                      := L      0.1,
           IN2                      := L      0.2,
           OUT3                     := M     19.2,
           OUT4                     := Q      0.0);
      NOP   0;
NETWORK
TITLE =

      A(    ;
      A     I    134.5;
      A(    ;
      O     M      4.1;
      O     M      4.2;
      )     ;
      O     ;
      A     I      1.6;
      A     M      4.0;
      )     ;
      AN    I      4.3;
      =     M     20.0;
NETWORK
TITLE =
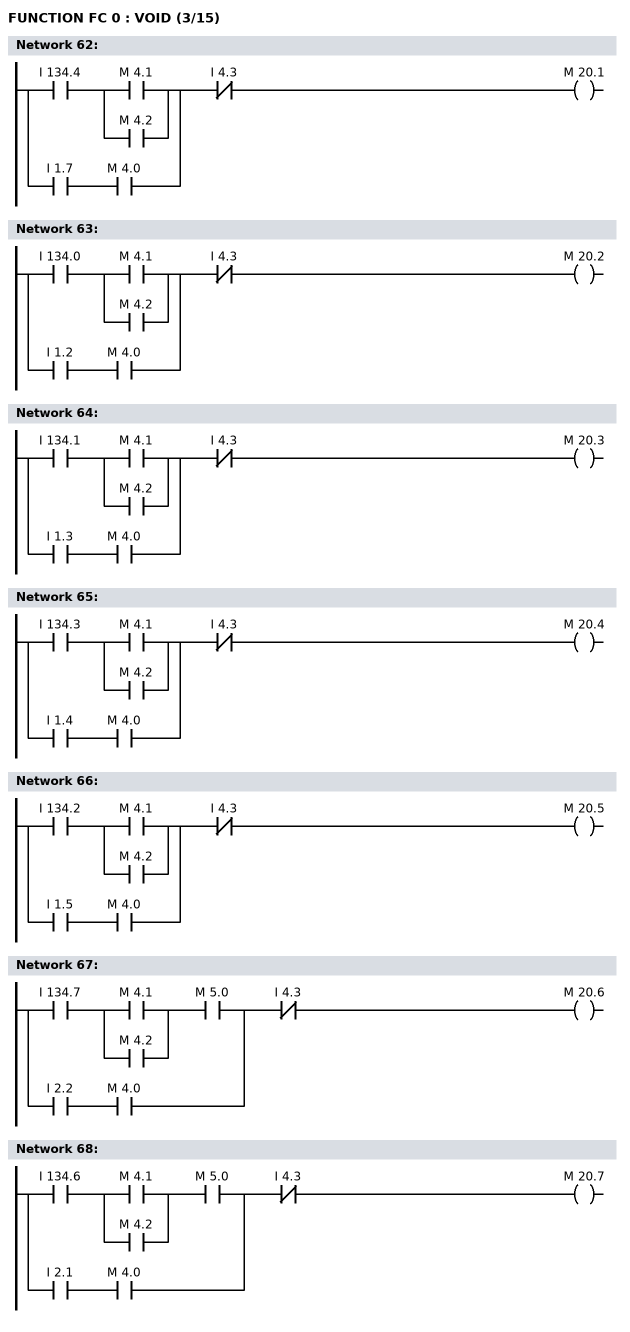

      A(    ;
      A     I    134.4;
      A(    ;
      O     M      4.1;
      O     M      4.2;
      )     ;
      O     ;
      A     I      1.7;
      A     M      4.0;
      )     ;
      AN    I      4.3;
      =     M     20.1;
NETWORK
TITLE =

      A(    ;
      A     I    134.0;
      A(    ;
      O     M      4.1;
      O     M      4.2;
      )     ;
      O     ;
      A     I      1.2;
      A     M      4.0;
      )     ;
      AN    I      4.3;
      =     M     20.2;
NETWORK
TITLE =

      A(    ;
      A     I    134.1;
      A(    ;
      O     M      4.1;
      O     M      4.2;
      )     ;
      O     ;
      A     I      1.3;
      A     M      4.0;
      )     ;
      AN    I      4.3;
      =     M     20.3;
NETWORK
TITLE =

      A(    ;
      A     I    134.3;
      A(    ;
      O     M      4.1;
      O     M      4.2;
      )     ;
      O     ;
      A     I      1.4;
      A     M      4.0;
      )     ;
      AN    I      4.3;
      =     M     20.4;
NETWORK
TITLE =

      A(    ;
      A     I    134.2;
      A(    ;
      O     M      4.1;
      O     M      4.2;
      )     ;
      O     ;
      A     I      1.5;
      A     M      4.0;
      )     ;
      AN    I      4.3;
      =     M     20.5;
NETWORK
TITLE =

      A(    ;
      A     I    134.7;
      A(    ;
      O     M      4.1;
      O     M      4.2;
      )     ;
      A     M      5.0;
      O     ;
      A     I      2.2;
      A     M      4.0;
      )     ;
      AN    I      4.3;
      =     M     20.6;
NETWORK
TITLE =

      A(    ;
      A     I    134.6;
      A(    ;
      O     M      4.1;
      O     M      4.2;
      )     ;
      A     M      5.0;
      O     ;
      A     I      2.1;
      A     M      4.0;
      )     ;
      AN    I      4.3;
      =     M     20.7;
NETWORK
TITLE =
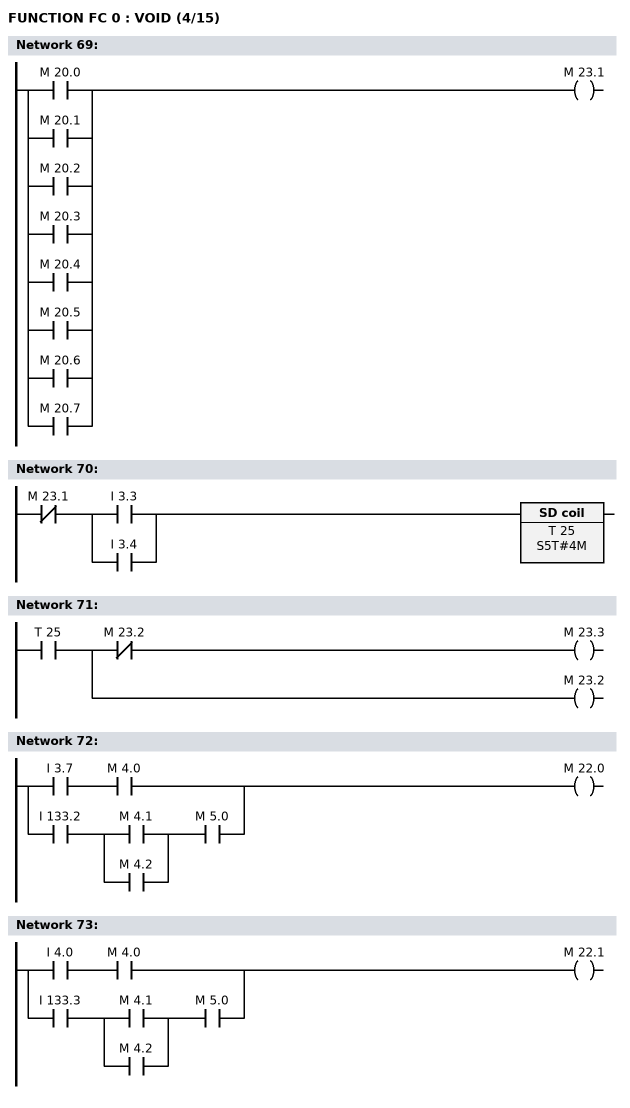

      O     M     20.0;
      O     M     20.1;
      O     M     20.2;
      O     M     20.3;
      O     M     20.4;
      O     M     20.5;
      O     M     20.6;
      O     M     20.7;
      =     M     23.1;
NETWORK
TITLE =

      AN    M     23.1;
      A(    ;
      O     I      3.3;
      O     I      3.4;
      )     ;
      L     S5T#4M;
      SD    T     25;
      NOP   0;
      NOP   0;
      NOP   0;
      NOP   0;
NETWORK
TITLE =

      A     T     25;
      =     L      0.0;
      A     L      0.0;
      AN    M     23.2;
      =     M     23.3;
      A     L      0.0;
      BLD   102;
      =     M     23.2;
NETWORK
TITLE =

      A     I      3.7;
      A     M      4.0;
      O     ;
      A     I    133.2;
      A(    ;
      O     M      4.1;
      O     M      4.2;
      )     ;
      A     M      5.0;
      =     M     22.0;
NETWORK
TITLE =

      A     I      4.0;
      A     M      4.0;
      O     ;
      A     I    133.3;
      A(    ;
      O     M      4.1;
      O     M      4.2;
      )     ;
      A     M      5.0;
      =     M     22.1;
NETWORK
TITLE =
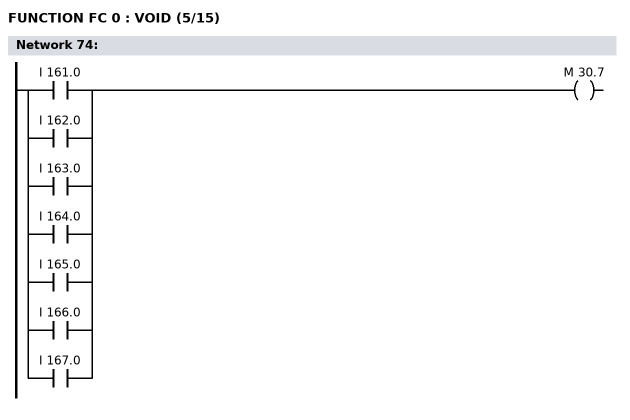

      O     I    161.0;
      O     I    162.0;
      O     I    163.0;
      O     I    164.0;
      O     I    165.0;
      O     I    166.0;
      O     I    167.0;
      =     M     30.7;
NETWORK
TITLE =
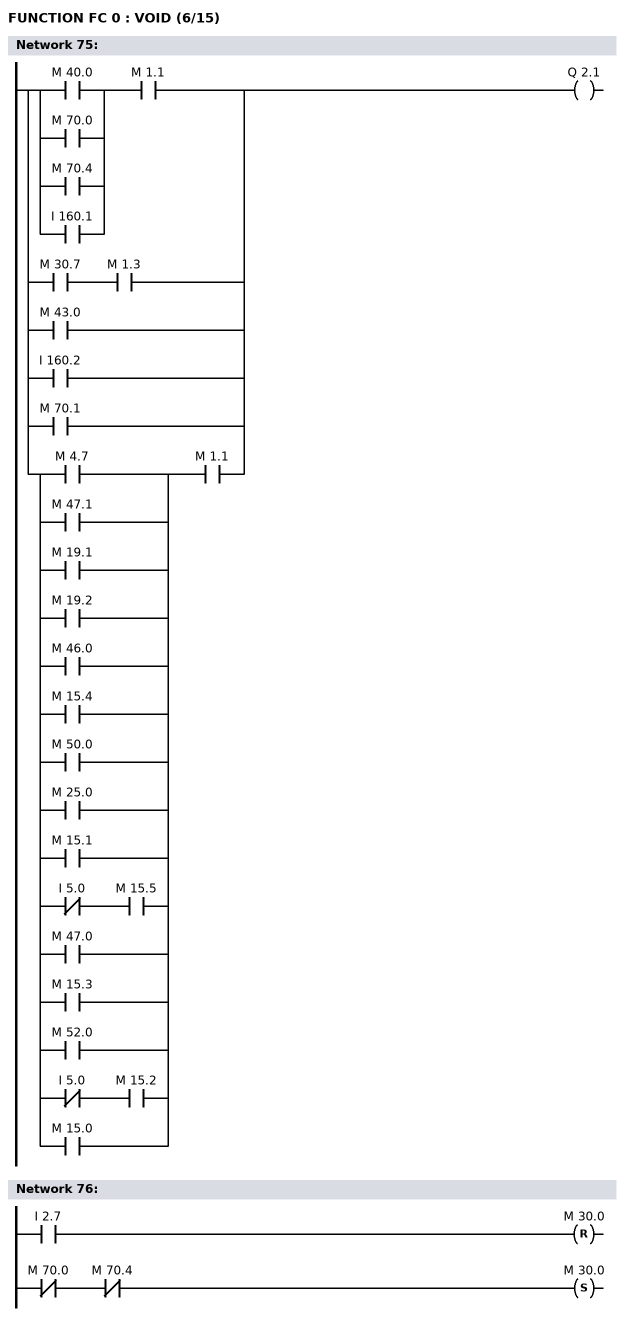

      A(    ;
      O     M     40.0;
      O     M     70.0;
      O     M     70.4;
      O     I    160.1;
      )     ;
      A     M      1.1;
      O     ;
      A     M     30.7;
      A     M      1.3;
      O     M     43.0;
      O     I    160.2;
      O     M     70.1;
      O     ;
      A(    ;
      O     M      4.7;
      O     M     47.1;
      O     M     19.1;
      O     M     19.2;
      O     M     46.0;
      O     M     15.4;
      O     M     50.0;
      O     M     25.0;
      O     M     15.1;
      O     ;
      AN    I      5.0;
      A     M     15.5;
      O     M     47.0;
      O     M     15.3;
      O     M     52.0;
      O     ;
      AN    I      5.0;
      A     M     15.2;
      O     M     15.0;
      )     ;
      A     M      1.1;
      =     Q      2.1;
NETWORK
TITLE =

      A     I      2.7;
      R     M     30.0;
      AN    M     70.0;
      AN    M     70.4;
      S     M     30.0;
      NOP   0;
NETWORK
TITLE =
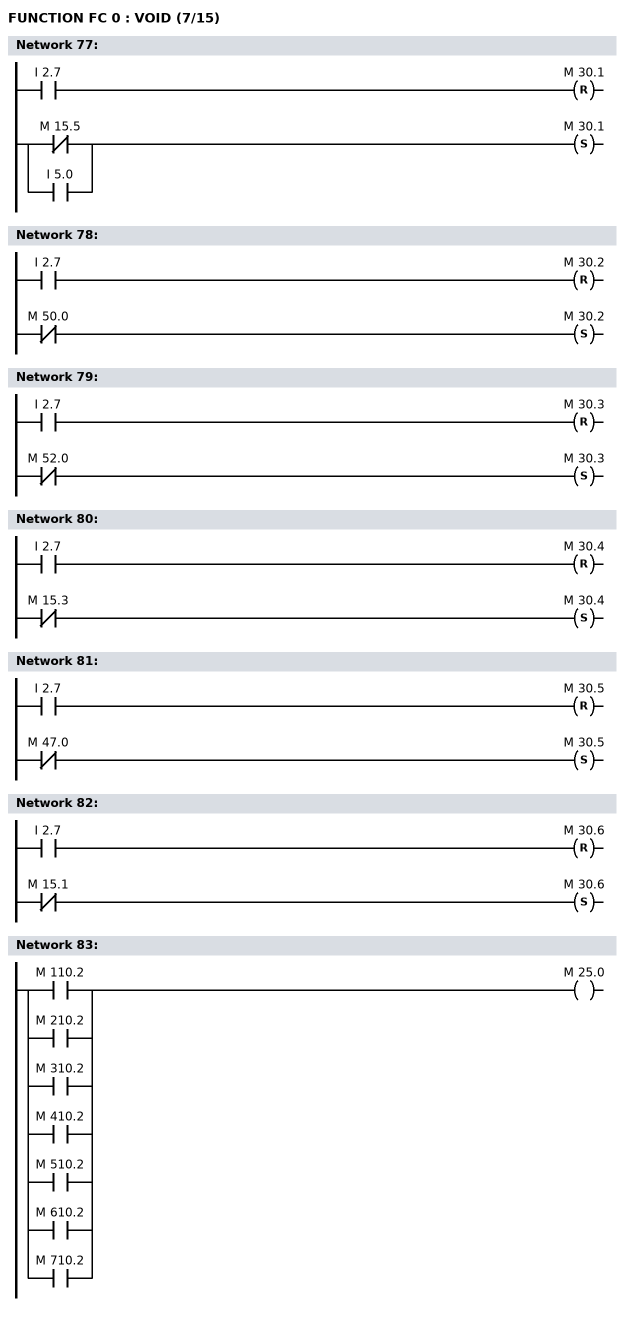

      A     I      2.7;
      R     M     30.1;
      A(    ;
      ON    M     15.5;
      O     I      5.0;
      )     ;
      S     M     30.1;
      NOP   0;
NETWORK
TITLE =

      A     I      2.7;
      R     M     30.2;
      AN    M     50.0;
      S     M     30.2;
      NOP   0;
NETWORK
TITLE =

      A     I      2.7;
      R     M     30.3;
      AN    M     52.0;
      S     M     30.3;
      NOP   0;
NETWORK
TITLE =

      A     I      2.7;
      R     M     30.4;
      AN    M     15.3;
      S     M     30.4;
      NOP   0;
NETWORK
TITLE =

      A     I      2.7;
      R     M     30.5;
      AN    M     47.0;
      S     M     30.5;
      NOP   0;
NETWORK
TITLE =

      A     I      2.7;
      R     M     30.6;
      AN    M     15.1;
      S     M     30.6;
      NOP   0;
NETWORK
TITLE =

      O     M    110.2;
      O     M    210.2;
      O     M    310.2;
      O     M    410.2;
      O     M    510.2;
      O     M    610.2;
      O     M    710.2;
      =     M     25.0;
NETWORK
TITLE =
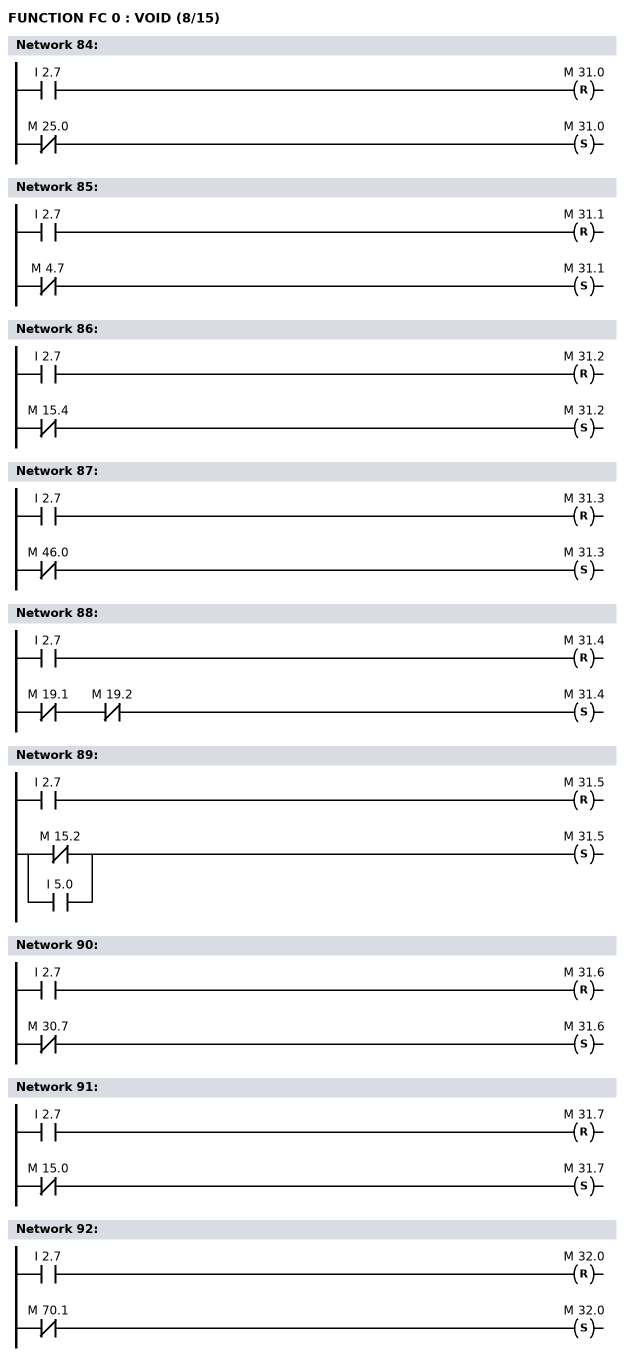

      A     I      2.7;
      R     M     31.0;
      AN    M     25.0;
      S     M     31.0;
      NOP   0;
NETWORK
TITLE =

      A     I      2.7;
      R     M     31.1;
      AN    M      4.7;
      S     M     31.1;
      NOP   0;
NETWORK
TITLE =

      A     I      2.7;
      R     M     31.2;
      AN    M     15.4;
      S     M     31.2;
      NOP   0;
NETWORK
TITLE =

      A     I      2.7;
      R     M     31.3;
      AN    M     46.0;
      S     M     31.3;
      NOP   0;
NETWORK
TITLE =

      A     I      2.7;
      R     M     31.4;
      AN    M     19.1;
      AN    M     19.2;
      S     M     31.4;
      NOP   0;
NETWORK
TITLE =

      A     I      2.7;
      R     M     31.5;
      A(    ;
      ON    M     15.2;
      O     I      5.0;
      )     ;
      S     M     31.5;
      NOP   0;
NETWORK
TITLE =

      A     I      2.7;
      R     M     31.6;
      AN    M     30.7;
      S     M     31.6;
      NOP   0;
NETWORK
TITLE =

      A     I      2.7;
      R     M     31.7;
      AN    M     15.0;
      S     M     31.7;
      NOP   0;
NETWORK
TITLE =

      A     I      2.7;
      R     M     32.0;
      AN    M     70.1;
      S     M     32.0;
      NOP   0;
NETWORK
TITLE =
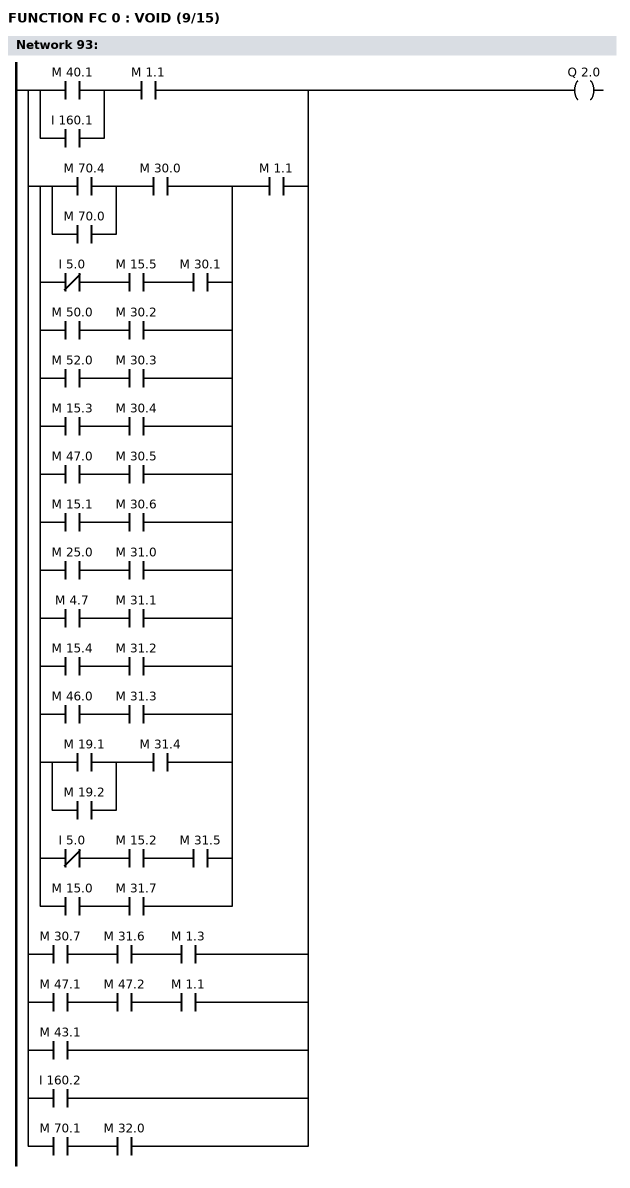

      A(    ;
      O     M     40.1;
      O     I    160.1;
      )     ;
      A     M      1.1;
      O     ;
      A(    ;
      A(    ;
      O     M     70.4;
      O     M     70.0;
      )     ;
      A     M     30.0;
      O     ;
      AN    I      5.0;
      A     M     15.5;
      A     M     30.1;
      O     ;
      A     M     50.0;
      A     M     30.2;
      O     ;
      A     M     52.0;
      A     M     30.3;
      O     ;
      A     M     15.3;
      A     M     30.4;
      O     ;
      A     M     47.0;
      A     M     30.5;
      O     ;
      A     M     15.1;
      A     M     30.6;
      O     ;
      A     M     25.0;
      A     M     31.0;
      O     ;
      A     M      4.7;
      A     M     31.1;
      O     ;
      A     M     15.4;
      A     M     31.2;
      O     ;
      A     M     46.0;
      A     M     31.3;
      O     ;
      A(    ;
      O     M     19.1;
      O     M     19.2;
      )     ;
      A     M     31.4;
      O     ;
      AN    I      5.0;
      A     M     15.2;
      A     M     31.5;
      O     ;
      A     M     15.0;
      A     M     31.7;
      )     ;
      A     M      1.1;
      O     ;
      A     M     30.7;
      A     M     31.6;
      A     M      1.3;
      O     ;
      A     M     47.1;
      A     M     47.2;
      A     M      1.1;
      O     M     43.1;
      O     I    160.2;
      O     ;
      A     M     70.1;
      A     M     32.0;
      =     Q      2.0;
NETWORK
TITLE =
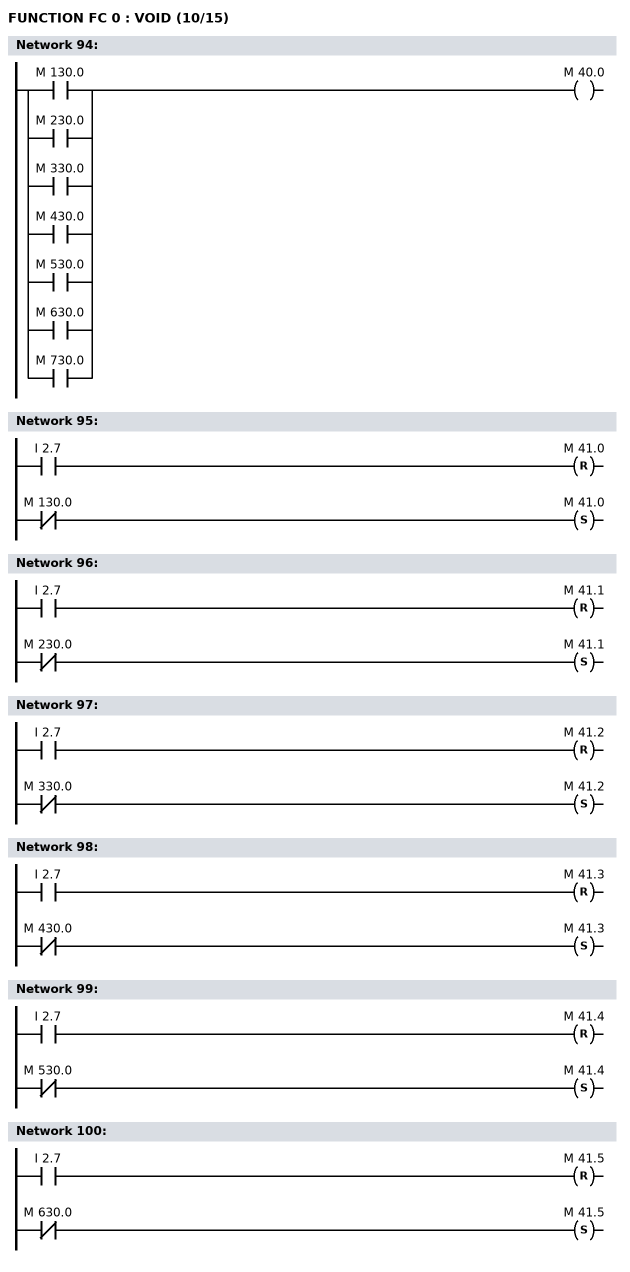

      O     M    130.0;
      O     M    230.0;
      O     M    330.0;
      O     M    430.0;
      O     M    530.0;
      O     M    630.0;
      O     M    730.0;
      =     M     40.0;
NETWORK
TITLE =

      A     I      2.7;
      R     M     41.0;
      AN    M    130.0;
      S     M     41.0;
      NOP   0;
NETWORK
TITLE =

      A     I      2.7;
      R     M     41.1;
      AN    M    230.0;
      S     M     41.1;
      NOP   0;
NETWORK
TITLE =

      A     I      2.7;
      R     M     41.2;
      AN    M    330.0;
      S     M     41.2;
      NOP   0;
NETWORK
TITLE =

      A     I      2.7;
      R     M     41.3;
      AN    M    430.0;
      S     M     41.3;
      NOP   0;
NETWORK
TITLE =

      A     I      2.7;
      R     M     41.4;
      AN    M    530.0;
      S     M     41.4;
      NOP   0;
NETWORK
TITLE =

      A     I      2.7;
      R     M     41.5;
      AN    M    630.0;
      S     M     41.5;
      NOP   0;
NETWORK
TITLE =
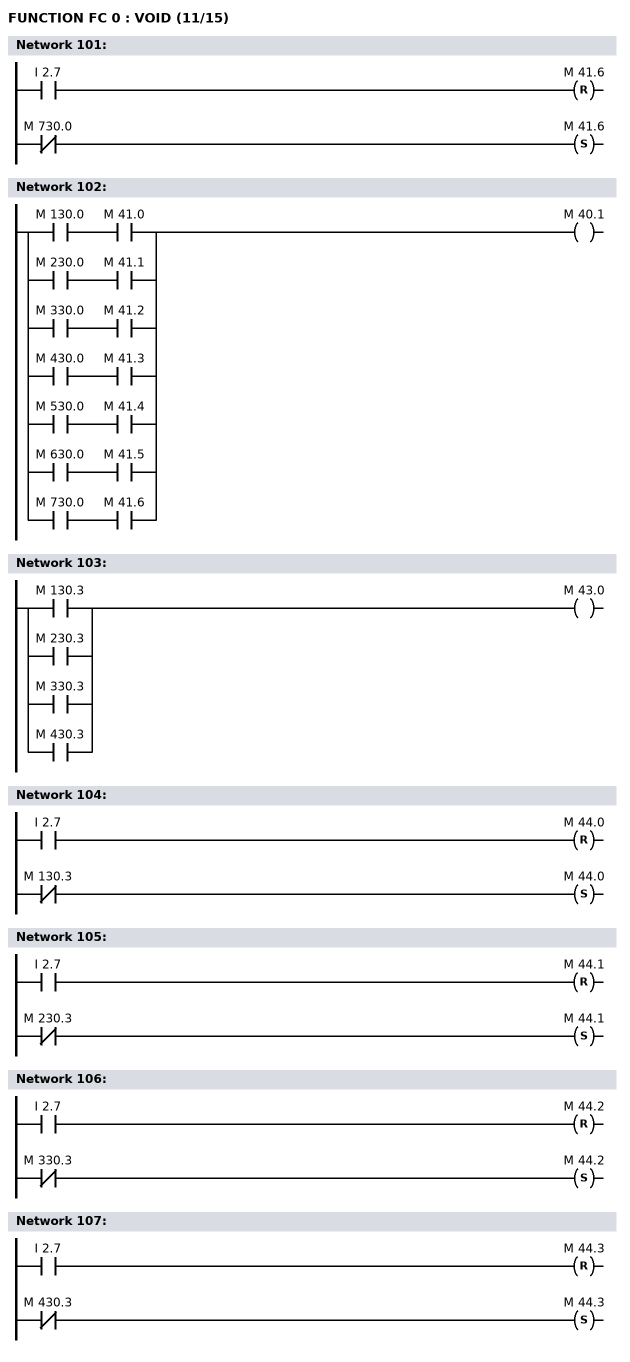

      A     I      2.7;
      R     M     41.6;
      AN    M    730.0;
      S     M     41.6;
      NOP   0;
NETWORK
TITLE =

      A     M    130.0;
      A     M     41.0;
      O     ;
      A     M    230.0;
      A     M     41.1;
      O     ;
      A     M    330.0;
      A     M     41.2;
      O     ;
      A     M    430.0;
      A     M     41.3;
      O     ;
      A     M    530.0;
      A     M     41.4;
      O     ;
      A     M    630.0;
      A     M     41.5;
      O     ;
      A     M    730.0;
      A     M     41.6;
      =     M     40.1;
NETWORK
TITLE =

      O     M    130.3;
      O     M    230.3;
      O     M    330.3;
      O     M    430.3;
      =     M     43.0;
NETWORK
TITLE =

      A     I      2.7;
      R     M     44.0;
      AN    M    130.3;
      S     M     44.0;
      NOP   0;
NETWORK
TITLE =

      A     I      2.7;
      R     M     44.1;
      AN    M    230.3;
      S     M     44.1;
      NOP   0;
NETWORK
TITLE =

      A     I      2.7;
      R     M     44.2;
      AN    M    330.3;
      S     M     44.2;
      NOP   0;
NETWORK
TITLE =

      A     I      2.7;
      R     M     44.3;
      AN    M    430.3;
      S     M     44.3;
      NOP   0;
NETWORK
TITLE =
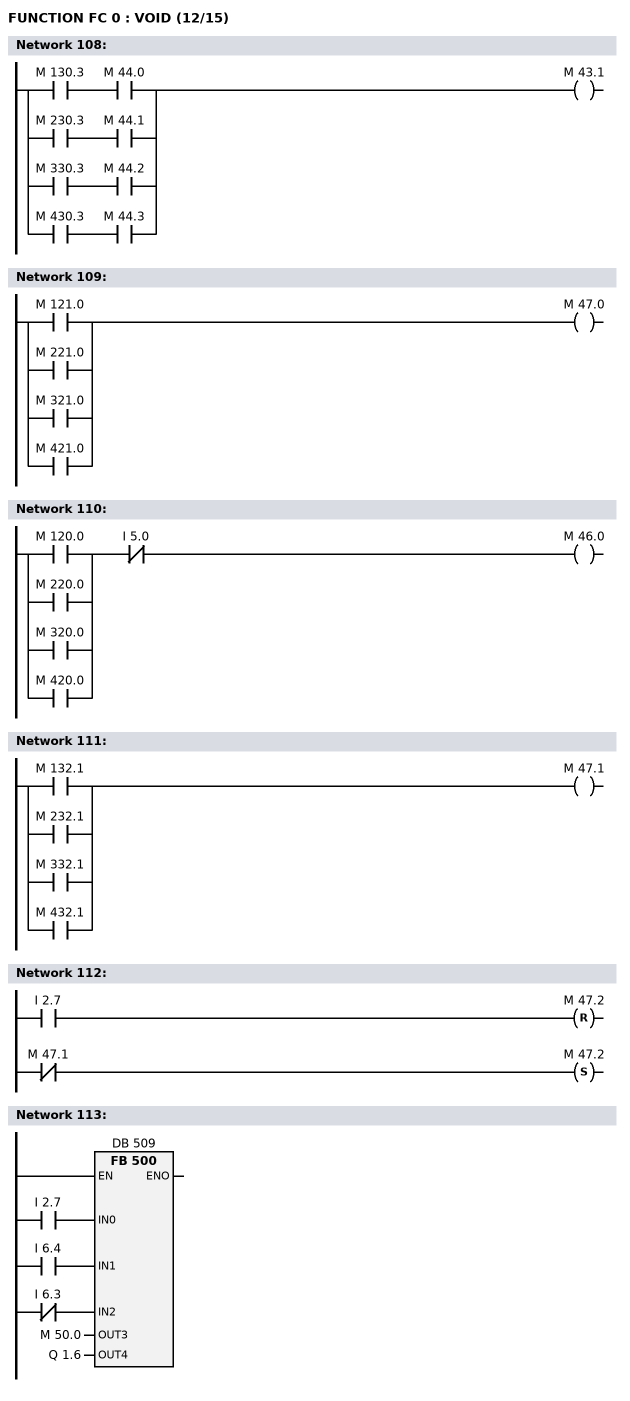

      A     M    130.3;
      A     M     44.0;
      O     ;
      A     M    230.3;
      A     M     44.1;
      O     ;
      A     M    330.3;
      A     M     44.2;
      O     ;
      A     M    430.3;
      A     M     44.3;
      =     M     43.1;
NETWORK
TITLE =

      O     M    121.0;
      O     M    221.0;
      O     M    321.0;
      O     M    421.0;
      =     M     47.0;
NETWORK
TITLE =

      A(    ;
      O     M    120.0;
      O     M    220.0;
      O     M    320.0;
      O     M    420.0;
      )     ;
      AN    I      5.0;
      =     M     46.0;
NETWORK
TITLE =

      O     M    132.1;
      O     M    232.1;
      O     M    332.1;
      O     M    432.1;
      =     M     47.1;
NETWORK
TITLE =

      A     I      2.7;
      R     M     47.2;
      AN    M     47.1;
      S     M     47.2;
      NOP   0;
NETWORK
TITLE =

      A     I      2.7;
      =     L      0.0;
      BLD   103;
      A     I      6.4;
      =     L      0.1;
      BLD   103;
      AN    I      6.3;
      =     L      0.2;
      BLD   103;
      CALL FB   500 , DB   509 (
           IN0                      := L      0.0,
           IN1                      := L      0.1,
           IN2                      := L      0.2,
           OUT3                     := M     50.0,
           OUT4                     := Q      1.6);
      NOP   0;
NETWORK
TITLE =
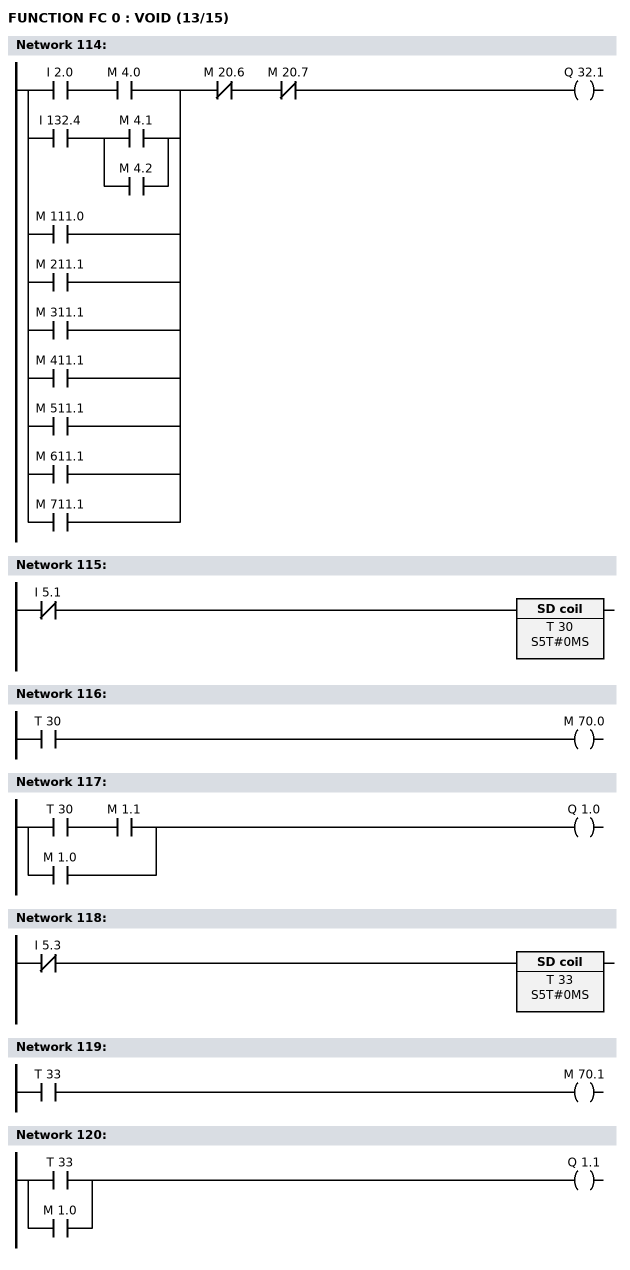

      A(    ;
      A     I      2.0;
      A     M      4.0;
      O     ;
      A     I    132.4;
      A(    ;
      O     M      4.1;
      O     M      4.2;
      )     ;
      O     M    111.0;
      O     M    211.1;
      O     M    311.1;
      O     M    411.1;
      O     M    511.1;
      O     M    611.1;
      O     M    711.1;
      )     ;
      AN    M     20.6;
      AN    M     20.7;
      =     Q     32.1;
NETWORK
TITLE =

      AN    I      5.1;
      L     S5T#0MS;
      SD    T     30;
      NOP   0;
      NOP   0;
      NOP   0;
      NOP   0;
NETWORK
TITLE =

      A     T     30;
      =     M     70.0;
NETWORK
TITLE =

      A     T     30;
      A     M      1.1;
      O     M      1.0;
      =     Q      1.0;
NETWORK
TITLE =

      AN    I      5.3;
      L     S5T#0MS;
      SD    T     33;
      NOP   0;
      NOP   0;
      NOP   0;
      NOP   0;
NETWORK
TITLE =

      A     T     33;
      =     M     70.1;
NETWORK
TITLE =

      O     T     33;
      O     M      1.0;
      =     Q      1.1;
NETWORK
TITLE =
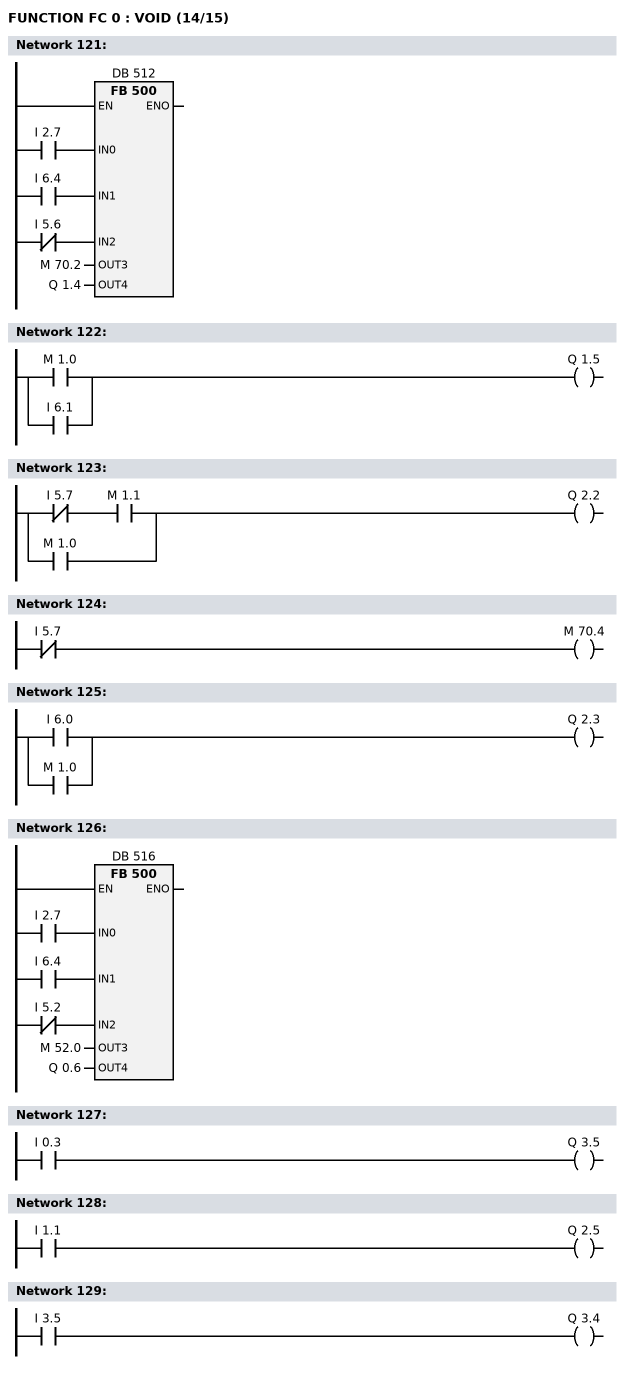

      A     I      2.7;
      =     L      0.0;
      BLD   103;
      A     I      6.4;
      =     L      0.1;
      BLD   103;
      AN    I      5.6;
      =     L      0.2;
      BLD   103;
      CALL FB   500 , DB   512 (
           IN0                      := L      0.0,
           IN1                      := L      0.1,
           IN2                      := L      0.2,
           OUT3                     := M     70.2,
           OUT4                     := Q      1.4);
      NOP   0;
NETWORK
TITLE =

      O     M      1.0;
      O     I      6.1;
      =     Q      1.5;
NETWORK
TITLE =

      AN    I      5.7;
      A     M      1.1;
      O     M      1.0;
      =     Q      2.2;
NETWORK
TITLE =

      AN    I      5.7;
      =     M     70.4;
NETWORK
TITLE =

      O     I      6.0;
      O     M      1.0;
      =     Q      2.3;
NETWORK
TITLE =

      A     I      2.7;
      =     L      0.0;
      BLD   103;
      A     I      6.4;
      =     L      0.1;
      BLD   103;
      AN    I      5.2;
      =     L      0.2;
      BLD   103;
      CALL FB   500 , DB   516 (
           IN0                      := L      0.0,
           IN1                      := L      0.1,
           IN2                      := L      0.2,
           OUT3                     := M     52.0,
           OUT4                     := Q      0.6);
      NOP   0;
NETWORK
TITLE =

      A     I      0.3;
      =     Q      3.5;
NETWORK
TITLE =

      A     I      1.1;
      =     Q      2.5;
NETWORK
TITLE =

      A     I      3.5;
      =     Q      3.4;
NETWORK
TITLE =
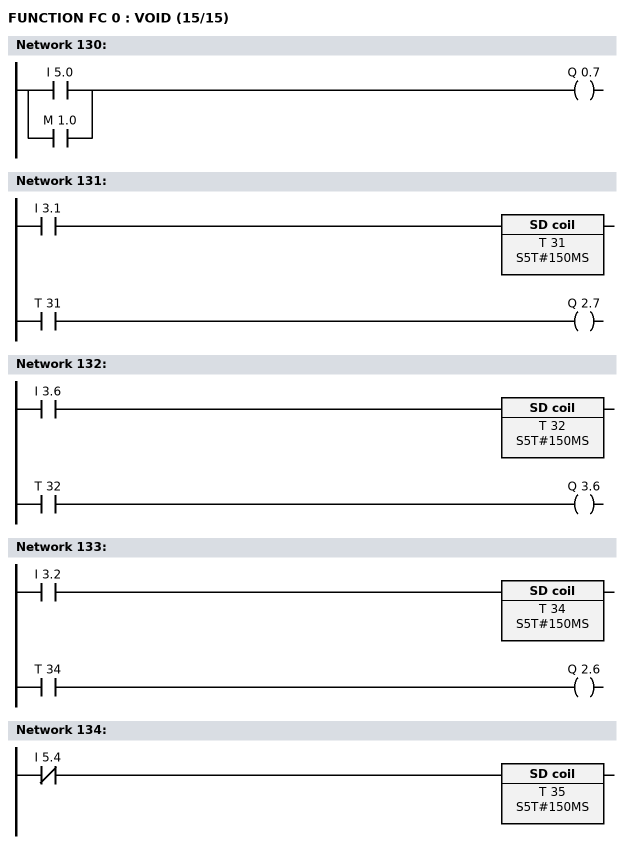

      O     I      5.0;
      O     M      1.0;
      =     Q      0.7;
NETWORK
TITLE =

      A     I      3.1;
      L     S5T#150MS;
      SD    T     31;
      NOP   0;
      NOP   0;
      NOP   0;
      A     T     31;
      =     Q      2.7;
NETWORK
TITLE =

      A     I      3.6;
      L     S5T#150MS;
      SD    T     32;
      NOP   0;
      NOP   0;
      NOP   0;
      A     T     32;
      =     Q      3.6;
NETWORK
TITLE =

      A     I      3.2;
      L     S5T#150MS;
      SD    T     34;
      NOP   0;
      NOP   0;
      NOP   0;
      A     T     34;
      =     Q      2.6;
NETWORK
TITLE =

      AN    I      5.4;
      L     S5T#150MS;
      SD    T     35;
      NOP   0;
      NOP   0;
      NOP   0;
      NOP   0;
END_FUNCTION

FUNCTION FC 1 : VOID
VERSION : 0.1

BEGIN
NETWORK
TITLE =
